         // Create log entry
         CreateLogMessagePara2 ( Timestamp   := SystemTime,
                                 MessageType := MessageType.CMD,
                                 Severity    := Severity.DEBUG,
                                 MessageCode := 0,
                                 MessageText := 'SyncSwLimits: Synchronization of SwLimits triggered by RC, SyncMode = {1}, SyncTime = {2}, SyncDirection = PLC -> RC',
                                 Para1       :=  SYNC_MODE_TO_STRING(AxesGroup.Parameter.Plc.Parameter.SynchronizationModes.SWLimits[SyncTime.AFTER_START_UP]),
                                 Para2       :=  SYNC_TIME_TO_STRING(SyncTime.AFTER_START_UP));
                                 RETURN;
			 END_IF
       
       // set timeout
       SetTimeout(PT := _rTimeout, rTimer := _rTimer);
       // jump back
      _rStep := 10;

       
  // ------------------------------------------
  // SyncMode : SERVER_TO_CLIENT 
  // ------------------------------------------
  12 : // Conflict triggerd by PLC ?  
       IF ( NOT AxesGroup.State.SyncStatePlc.InSync.SwLimits )
       THEN
         // set timeout
         SetTimeout(PT := _rTimeout, rTimer := _rTimer);
         // inc step counter
        _rStep := 20; // -> read RC data and write it to PLC                  

         // Create log entry
         CreateLogMessagePara2 ( Timestamp   := SystemTime,
                                 MessageType := MessageType.CMD,
                                 Severity    := Severity.DEBUG,
                                 MessageCode := 0,
                                 MessageText := 'SyncSwLimits: Synchronization of SwLimits triggered by PLC, SyncMode = {1}, SyncTime = {2}, SyncDirection = RC -> PLC',
                                 Para1       :=  SYNC_MODE_TO_STRING(AxesGroup.Parameter.Plc.Parameter.SynchronizationModes.SWLimits[SyncTime.AFTER_START_UP]),
                                 Para2       :=  SYNC_TIME_TO_STRING(SyncTime.AFTER_START_UP));
                                 RETURN;
       END_IF
   
       // Conflict triggered by RC ?
       IF ( NOT AxesGroup.State.SyncStateRc.InSync.SwLimits )
       THEN
         // set timeout
         SetTimeout(PT := _rTimeout, rTimer := _rTimer);
         // inc step counter
        _rStep := 20; // -> read RC data and write it to PLC

         // Create log entry
         CreateLogMessagePara2 ( Timestamp   := SystemTime,
                                 MessageType := MessageType.CMD,
                                 Severity    := Severity.DEBUG,
                                 MessageCode := 0,
                                 MessageText := 'SyncSwLimits: Synchronization of SwLimits triggered by RC, SyncMode = {1}, SyncTime = {2}, SyncDirection = RC -> PLC',
                                 Para1       :=  SYNC_MODE_TO_STRING(AxesGroup.Parameter.Plc.Parameter.SynchronizationModes.SWLimits[SyncTime.AFTER_START_UP]),
                                 Para2       :=  SYNC_TIME_TO_STRING(SyncTime.AFTER_START_UP));
                                 RETURN;
			 END_IF
       
       // set timeout
       SetTimeout(PT := _rTimeout, rTimer := _rTimer);
       // jump back
      _rStep := 10;
  

  // ------------------------------------------
  // SyncMode : AUTOMATIC 
  // ------------------------------------------
  13 : // Conflict triggerd by PLC ?  
       IF ( NOT AxesGroup.State.SyncStatePlc.InSync.SwLimits )
       THEN
         // set timeout
         SetTimeout(PT := _rTimeout, rTimer := _rTimer);
         // inc step counter
        _rStep := 30; // -> write PLC data to RC                  
         
         // Create log entry
         CreateLogMessagePara2 ( Timestamp   := SystemTime,
                                 MessageType := MessageType.CMD,
                                 Severity    := Severity.DEBUG,
                                 MessageCode := 0,
                                 MessageText := 'SyncSwLimits: Synchronization of SwLimits triggered by PLC, SyncMode = {1}, SyncTime = {2}, SyncDirection = PLC -> RC',
                                 Para1       :=  SYNC_MODE_TO_STRING(AxesGroup.Parameter.Plc.Parameter.SynchronizationModes.SWLimits[SyncTime.AFTER_START_UP]),
                                 Para2       :=  SYNC_TIME_TO_STRING(SyncTime.AFTER_START_UP));
                                 RETURN;
       END_IF
   
       // Conflict triggered by RC ?
       IF ( NOT AxesGroup.State.SyncStateRc.InSync.SwLimits )
       THEN
         // set timeout
         SetTimeout(PT := _rTimeout, rTimer := _rTimer);
         // inc step counter
        _rStep := 20; // -> read RC data an write it to PLC

         // Create log entry
         CreateLogMessagePara2 ( Timestamp   := SystemTime,
                                 MessageType := MessageType.CMD,
                                 Severity    := Severity.DEBUG,
                                 MessageCode := 0,
                                 MessageText := 'SyncSwLimits: Synchronization of SwLimits triggered by RC, SyncMode = {1}, SyncTime = {2}, SyncDirection = RC -> PLC',
                                 Para1       :=  SYNC_MODE_TO_STRING(AxesGroup.Parameter.Plc.Parameter.SynchronizationModes.SWLimits[SyncTime.AFTER_START_UP]),
                                 Para2       :=  SYNC_TIME_TO_STRING(SyncTime.AFTER_START_UP));
                                 RETURN;
			 END_IF
       
       // set timeout
       SetTimeout(PT := _rTimeout, rTimer := _rTimer);
       // jump back
      _rStep := 10; // ST-FIX F95: was commented out


  // ------------------------------------------
  // Read Data from RC and write it to PLC
  // ------------------------------------------
  20 : IF (( NOT _readRobotSWLimits.Busy  ) AND 
           ( NOT _readRobotSWLimits.Error ))
       THEN
         // execute command
        _readRobotSWLimits.Execute := TRUE;
         // set timeout
         SetTimeout(PT := _rTimeout, rTimer := _rTimer);
         // inc step counter
        _rStep := _rStep + 1;
       ELSE
         // check error ? 
         IF (_readRobotSWLimits.Error)
         THEN
           ErrorID     := _readRobotSWLimits.ErrorID;
           ErrorAddTxt := _readRobotSWLimits.ErrorAddTxt;
         END_IF  
       
         // timeout exceeded ? 
         IF (CheckTimeout(_rTimer) = RobotLibraryConstants.OK)
         THEN
           ErrorID     := RobotLibraryErrorIdEnum.ERR_TIMEOUT_CMD;
           ErrorAddTxt := CONCAT(_stepName, DINT_TO_STRING(_rStep));
         END_IF
       END_IF
 
  21 : IF (( NOT _readRobotSWLimits.Busy  ) AND
           ( NOT _readRobotSWLimits.Error ) AND
           (     _readRobotSWLimits.Done  ))
       THEN
         // reset execution
        _readRobotSWLimits.Execute := FALSE;
         // ST-FIX F107: AUTOMATIC - the PLC data were changed while the RC data were read: the PLC
         // change is the most recent one and is written to the RC instead of being overwritten
         IF ( AxesGroup.Parameter.Plc.Parameter.SynchronizationModes.SWLimits[SyncTime.AFTER_START_UP] = SyncMode.AUTOMATIC ) AND
            ( NOT IsSwLimitsEqual( Data1 := SwLimits, Data2 := _swLimits, IgnoreTimestamp := TRUE ))
         THEN
           // set timeout
           SetTimeout(PT := _rTimeout, rTimer := _rTimer);
           // -> write PLC data to RC
          _rStep := 30;
           RETURN;
         END_IF
         // update internal SwLimits data
         SwLimits := _readRobotSWLimits.OutCmd.LimitValues;         
        _swLimits := _readRobotSWLimits.OutCmd.LimitValues;
         // set timeout
         SetTimeout(PT := _rTimeout, rTimer := _rTimer);
         // inc step counter
        // ST-FIX F20: write the RC data back to reset DataChanged on the RC (spec 5.6.7.4.2)
        IF ( AxesGroup.State.RobotData.RCSupportedFunctions.WriteRobotSWLimits )
        THEN
          _rStep := 30;
        ELSE
          _rStep := 10;
        END_IF // -> jump to after startup           
       ELSE
         // check error ? 
         IF (_readRobotSWLimits.Error)
         THEN
           ErrorID     := _readRobotSWLimits.ErrorID;
           ErrorAddTxt := _readRobotSWLimits.ErrorAddTxt;           
         END_IF  
       
         // timeout exceeded ? 
         IF (CheckTimeout(_rTimer) = RobotLibraryConstants.OK)
         THEN
           ErrorID     := RobotLibraryErrorIdEnum.ERR_TIMEOUT_CMD;
           ErrorAddTxt := CONCAT(_stepName, DINT_TO_STRING(_rStep));
         END_IF
       END_IF


  // ------------------------------------------
  // Write data from PLC to RC
  // ------------------------------------------
  30 : IF (( NOT _writeRobotSWLimits.Busy  ) AND 
           ( NOT _writeRobotSWLimits.Error ))
       THEN
         // set command parameter
        _writeRobotSWLimits.ParCmd.ResetToFactoryDefaults := FALSE;      
        _writeRobotSWLimits.ParCmd.LimitValues :=  SwLimits;
         // execute command
        _writeRobotSWLimits.Execute := TRUE;
         // set timeout
         SetTimeout(PT := _rTimeout, rTimer := _rTimer);
         // inc step counter
        _rStep := _rStep + 1;
       ELSE
         // check error ? 
         IF (_writeRobotSWLimits.Error)
         THEN
           ErrorID     := _writeRobotSWLimits.ErrorID;
           ErrorAddTxt := _writeRobotSWLimits.ErrorAddTxt;;
         END_IF  
       
         // timeout exceeded ? 
         IF (CheckTimeout(_rTimer) = RobotLibraryConstants.OK)
         THEN
           ErrorID     := RobotLibraryErrorIdEnum.ERR_TIMEOUT_CMD;
           ErrorAddTxt := CONCAT(_stepName, DINT_TO_STRING(_rStep));
         END_IF
       END_IF
 
  31 : IF (( NOT _writeRobotSWLimits.Busy  ) AND
           ( NOT _writeRobotSWLimits.Error ) AND
           (     _writeRobotSWLimits.Done  ))
       THEN
         // execute command
        _writeRobotSWLimits.Execute := FALSE;      
         // update internal SwLimits data
        _swLimits := SwLimits; 
         // set timeout
         SetTimeout(PT := _rTimeout, rTimer := _rTimer);
         // inc step counter
        _rStep := 10; // -> jump to after startup;           
       ELSE
         // check error ? 
         IF (_writeRobotSWLimits.Error)
         THEN
           SetWarning( WarningID := RobotLibraryWarningIdEnum.WARN_SW_LIMITS_SYNC_FAILED_BY_ERROR_OF_READ_OR_WRITE_CMD, Overwrite := TRUE);    
         END_IF  
       
         // timeout exceeded ? 
         IF (CheckTimeout(_rTimer) = RobotLibraryConstants.OK)
         THEN
           ErrorID     := RobotLibraryErrorIdEnum.ERR_TIMEOUT_CMD;
           ErrorAddTxt := CONCAT(_stepName, DINT_TO_STRING(_rStep));
         END_IF
       END_IF
       
ELSE
  // invalid step
  ErrorID     := RobotLibraryErrorIdEnum.ERR_INVALID_STEP;
  ErrorAddTxt := CONCAT(_stepName , DINT_TO_STRING(_stepCmd));
END_CASE
END_METHOD

METHOD PRIVATE HandleSyncToolData
VAR_IN_OUT
   /// Robot assignment of function
  AxesGroup : AxesGroup;
  /// ToolData stored on PLC.For more information refer to 5.5.6.4
  ToolData  : ARRAY[*] OF Tool;
END_VAR 

VAR
  /// Internal step counter name
 _stepName        : STRING;    
  /// Internal reference to step counter
 _rStep           : REFERENCE TO DINT;
  /// Internal reference to timer
 _rTimer          : REFERENCE TO TON;
  /// Internal reference to timeout
 _rTimeout        : REFERENCE TO TIME; 
  /// Internal reference to synchroniztion index
 _rSyncIdx        : REFERENCE TO USINT;
  /// internal bit for condition found
 _found           : BOOL;
  /// empty data set to reset all DataChanged bits
 _dataChangedNone : AxesGroupStateDataChanged; 
  /// internal index for loops
 _idx             : DINT;
END_VAR
// Set internal references 
_stepName      :=   '_stepSyncToolData = ';
_rStep       REF=    _stepSyncToolData;
_rTimer      REF=   _timerSyncToolData;
_rTimeout    REF= _timeoutSyncToolData;
_rSyncIdx    REF=     _syncIdxToolData;


CASE _rStep
OF    
  0: // Check initialisation configured ?
     // ST-FIX F130: an invalid sync mode (warning of CheckParameterValid) -> no synchronization of the data set
     IF ((( _parCfg.PLC.Parameter.SynchronizationModes.Tool[SyncTime.DURING_START_UP] = SyncMode.NO_SYNCHRONIZATION ) AND
          ( _parCfg.PLC.Parameter.SynchronizationModes.Tool[SyncTime. AFTER_START_UP] = SyncMode.NO_SYNCHRONIZATION )) OR
         ( NOT SyncModesValid( During := _parCfg.PLC.Parameter.SynchronizationModes.Tool[SyncTime.DURING_START_UP],
                               After  := _parCfg.PLC.Parameter.SynchronizationModes.Tool[SyncTime. AFTER_START_UP] ) ))
     THEN
       RETURN;
     END_IF
     

     // wait for initialisation done
     IF  ((     AxesGroup.State.RobotData.RCSupportedFunctions. ReadToolData ) AND
          (     AxesGroup.State.RobotData.RCSupportedFunctions.WriteToolData ) AND
          (     AxesGroup.State.Initialized                                  ) AND 
          ( NOT Error                                                        ))  
     THEN
       // ST-FIX F102: count check after the initialization (HighestXIndex of this connection)
     // Check More Data on RC than on PLC -> Synchronization not possible
     IF (AxesGroup.State.ConfigurationData.HighestToolIndex > AxesGroup.SystemData.ToolDataCount)
     THEN
       SetError( ErrorID := RobotLibraryErrorIdEnum.ERR_SYNC_TOOL_COUNT_RC_HIGHER_THAN_PLC, Overwrite := FALSE);
       RETURN;
		 END_IF
       // Check PLC tools < RC tools and SyncTool enabled ?    
       IF (( AxesGroup.State.DataEnableSync.EnableSyncTool      = TRUE                             )  AND
           ( AxesGroup.Parameter.Rob.Parameter.HighestToolIndex > AxesGroup.SystemData.ToolDataMax ))        
       THEN
         SetWarning( WarningID := RobotLibraryWarningIdEnum.WARN_TOOL_DATA_ARRAY_TOO_SHORT, Overwrite := TRUE);
       END_IF

       // Create log entry
       CreateLogMessagePara1 ( Timestamp   := SystemTime,
                               MessageType := MessageType.CMD,
                               Severity    := Severity.DEBUG,
                               MessageCode := 0,
                               MessageText := 'SyncToolData: Start initial reading of ToolData from RC',
                               Para1       :=  '');
       
       // init tool number
      _rSyncIdx := LIMIT(1, DINT_TO_USINT(AxesGroup.SystemData.ToolDataMin), AxesGroup.State.UnifiedToolIndex); // ST-FIX F21: index 0 is fixed on the RC 
       // init count of unsynchronized elements
       AxesGroup.State.SyncStatePlc.UnSyncNo.Tool := 0;
       // set timeout
       SetTimeout(PT := _rTimeout, rTimer := _rTimer);
       // inc step counter
      _rStep := _rStep + 1;
     END_IF     

     
     // Start read ToolData
  1: IF (( NOT _readToolData.Busy  ) AND 
         ( NOT _readToolData.Error ) AND
         ( NOT _readToolData.Done  ))
     THEN
       // set command parameter
      _readToolData.ParCmd.ToolNo := _rSyncIdx;      
       // execute command
      _readToolData.Execute := TRUE;
       // set timeout
       SetTimeout(PT := _rTimeout, rTimer := _rTimer);
       // inc step counter
      _rStep := _rStep + 1;
     ELSE
       // check error ? 
       IF ( _readToolData.Error ) AND ( WarningID = RobotLibraryWarningIdEnum.NO_WARNING )
       THEN
         SetWarning( WarningID := RobotLibraryWarningIdEnum.WARN_TOOL_SYNC_FAILED_BY_ERROR_OF_READ_OR_WRITE_CMD, Overwrite := TRUE);           
       END_IF  
       
       // timeout exceeded ? 
       IF (CheckTimeout(_rTimer) = RobotLibraryConstants.OK)
       THEN
         ErrorID     := RobotLibraryErrorIdEnum.ERR_TIMEOUT_CMD;
         ErrorAddTxt := CONCAT(_stepName, DINT_TO_STRING(_rStep));
       END_IF
     END_IF
 
     
     // Wait Tooldata read
  2: IF (( NOT _readToolData.Busy  ) AND
         ( NOT _readToolData.Error ) AND
         (     _readToolData.Done  ))
     THEN
       // reset execution
      _readToolData.Execute := FALSE;
       // set available bit
      _toolData[_rSyncIdx].Available := TRUE; 
       ToolData[_rSyncIdx].Available := TRUE;      
       // Copy data
      _toolData[_rSyncIdx].Data := _readToolData.OutCmd.ToolData;

       // Check tool data is equal ? 
       IF ( NOT IsToolDataEqual( Data1 := _toolData[_rSyncIdx].Data, Data2 := ToolData[_rSyncIdx].Data, IgnoreTimestamp := TRUE))
       THEN
         // Reset plc in sync flag
         AxesGroup.State.SyncStatePlc.InSync.Tool := FALSE;
         // Set data changed flag
         AxesGroup.State.DataChanged.Tool[_rSyncIdx] := TRUE;
         // inc count of unsynchronised plc tools
         AxesGroup.State.SyncStatePlc.UnSyncNo.Tool := AxesGroup.State.SyncStatePlc.UnSyncNo.Tool + 1;
        
         // Create log entry
         CreateLogMessagePara1 ( Timestamp   := SystemTime,
                                 MessageType := MessageType.CMD,
                                 Severity    := Severity.DEBUG,
                                 MessageCode := 0,
                                 MessageText := 'SyncToolData: Detected a difference in Tool[{1}] between PLC and RC',
                                 Para1       :=  DINT_TO_STRING(_rSyncIdx));
        
        
         // Check synchronisation is enabled ? 
         IF ( NOT AxesGroup.State.DataEnableSync.EnableSyncTool ) AND (InfoID = RobotLibraryInfoIdEnum.NO_INFO )
         THEN
           SetInfo( InfoID := RobotLibraryInfoIdEnum.INFO_SYNC_TOOL_DATA_DISABLED, Overwrite := TRUE);
				 END_IF
         
         // Check user interaction needed ?  
         IF ( AxesGroup.Parameter.PLC.Parameter.SyncUserInteraction.Tool ) AND ( WarningID = RobotLibraryWarningIdEnum.NO_WARNING )
         THEN
           SetWarning( WarningID := RobotLibraryWarningIdEnum.WARN_TOOL_NUMBER_SYNC_ERROR, Overwrite :=  TRUE);                    
				 END_IF
			 END_IF
             
       // Check all tools read ? 
       IF ( _rSyncIdx < AxesGroup.State.UnifiedToolIndex )
       THEN
         // set timeout
         SetTimeout(PT := _rTimeout, rTimer := _rTimer);
         // inc tool index
        _rSyncIdx := _rSyncIdx + 1;
         // dec step counter
        _rStep := _rStep - 1;
       ELSE
         // set timeout
         SetTimeout(PT := _rTimeout, rTimer := _rTimer);
         // inc step counter
        _rStep := _rStep + 1;           
       END_IF
     ELSE
       // check error ? 
       IF (_readToolData.Error)
       THEN
         // Set warning
         SetWarning( WarningID := RobotLibraryWarningIdEnum.WARN_TOOL_SYNC_FAILED_BY_ERROR_OF_READ_OR_WRITE_CMD, Overwrite := TRUE);                    
         // reset available bit
         ToolData[_rSyncIdx].Available := FALSE;
        _toolData[_rSyncIdx].Available := FALSE;
       END_IF  
       
       // timeout exceeded ? 
       IF (CheckTimeout(_rTimer) = RobotLibraryConstants.OK)
       THEN
         ErrorID     := RobotLibraryErrorIdEnum.ERR_TIMEOUT_CMD;
         ErrorAddTxt := CONCAT(_stepName, DINT_TO_STRING(_rStep));
       END_IF
     END_IF
     
     
     // Check synchronisation state ? 
  3: IF (( AxesGroup.State.SyncStatePlc.UnSyncNo.Tool                                            = 0                           ) OR 
         ( AxesGroup.Parameter.Plc.Parameter.SynchronizationModes.Tool[SyncTime.DURING_START_UP] = SyncMode.NO_SYNCHRONIZATION ))
     THEN
       // Update bit for data in sync
       AxesGroup.State.SyncStatePlc.InSync.Tool := (AxesGroup.State.SyncStatePlc.UnSyncNo.Tool = 0);
         // ST-FIX F165: synchronization of the start-up phase finished
         AxesGroup.State.Synchronizing.Tool := FALSE;
       // set timeout
       SetTimeout(PT := _rTimeout, rTimer := _rTimer);
       // inc step counter
      _rStep := 10; // -> jump to after startup
            
       // Create log entry
       CreateLogMessagePara1 ( Timestamp   := SystemTime,
                               MessageType := MessageType.CMD,
                               Severity    := Severity.DEBUG,
                               MessageCode := 0,
                               MessageText := 'SyncToolData: Synchronization Startup Phase done',
                               Para1       :=  '' );      
     ELSE 
       // Check user interaction needed ? 
       IF ( NOT AxesGroup.Parameter.PLC.Parameter.SyncUserInteraction.Tool )
       THEN
         CASE AxesGroup.Parameter.Plc.Parameter.SynchronizationModes.Tool[SyncTime.DURING_START_UP] OF

           SyncMode.SERVER_TO_CLIENT : 

           
             FOR _idx := AxesGroup.SystemData.ToolDataMin TO MIN(AxesGroup.SystemData.ToolDataMax, RobotLibraryParameter.TOOL_MAX - 1) // ST-FIX F18
             DO
               // Overwrite PLC data with RC data
               ToolData[_idx] := _toolData[_idx];            
						 END_FOR
             // Reset data changed flags
             AxesGroup.State.DataChanged.Tool := _dataChangedNone.Tool;
             // Reset Synchronizing flag
             AxesGroup.State.Synchronizing.Tool := FALSE;
             // Set plc in sync flag
             AxesGroup.State.SyncStatePlc.InSync.Tool := TRUE;
             // Reset count of unsynchronised plc tools
             AxesGroup.State.SyncStatePlc.UnSyncNo.Tool := 0;            
             // set timeout
             SetTimeout(PT := _rTimeout, rTimer := _rTimer);
             // inc step counter
            _rStep := 10; // -> jump to after startup         

            // Create log entry
            CreateLogMessagePara3 ( Timestamp   := SystemTime,
                                    MessageType := MessageType.CMD,
                                    Severity    := Severity.DEBUG,
                                    MessageCode := 0,
                                    MessageText := 'SyncToolData: Synchronization of Tools triggered by StartUp-Compare, SyncMode = {2}, SyncTime = {3}, SyncDirection = RC -> PLC',
                                    Para1       :=  DINT_TO_STRING(_rSyncIdx),
                                    Para2       :=  SYNC_MODE_TO_STRING(AxesGroup.Parameter.Plc.Parameter.SynchronizationModes.Tool[SyncTime.DURING_START_UP]),
                                    Para3       :=  SYNC_TIME_TO_STRING(SyncTime.DURING_START_UP));
            // Create log entry
            CreateLogMessagePara1 ( Timestamp   := SystemTime,
                                    MessageType := MessageType.CMD,
                                    Severity    := Severity.DEBUG,
                                    MessageCode := 0,
                                    MessageText := 'SyncToolData: Applied the initial read tool data from RC',
                                    Para1       :=  '' );

				   SyncMode.CLIENT_TO_SERVER : ;

             // Check conflicts to solve ? 
             FOR _rSyncIdx := 1 TO AxesGroup.State.UnifiedToolIndex // ST-FIX F21: index 0 is fixed on the RC
             DO
               IF ( AxesGroup.State.DataChanged.Tool[_rSyncIdx] )
               THEN
                _found := TRUE;
                 EXIT;
		  			   END_IF
             END_FOR
           
             IF ( _found ) 
             THEN
               // Reset plc in sync flag
               AxesGroup.State.SyncStatePlc.InSync.Tool := FALSE;
               // Set Synchronizing flag
               AxesGroup.State.Synchronizing.Tool := TRUE;
               // set timeout
               SetTimeout(PT := _rTimeout, rTimer := _rTimer);
               // inc step counter
              _rStep := _rStep +1; // -> write PLC data to RC                  
               // Create log entry
               CreateLogMessagePara3 ( Timestamp   := SystemTime,
                                       MessageType := MessageType.CMD,
                                       Severity    := Severity.DEBUG,
                                       MessageCode := 0,
                                       MessageText := 'SyncToolData: Synchronization of Tool[{1}] triggered by StartUp-Compare, SyncMode = {2}, SyncTime = {3}, SyncDirection = PLC -> RC',
                                       Para1       :=  DINT_TO_STRING(_rSyncIdx),
                                       Para2       :=  SYNC_MODE_TO_STRING(AxesGroup.Parameter.Plc.Parameter.SynchronizationModes.Tool[SyncTime.DURING_START_UP]),
                                       Para3       :=  SYNC_TIME_TO_STRING(SyncTime.DURING_START_UP));
             ELSE
               // Reset data changed flags
               AxesGroup.State.DataChanged.Tool := _dataChangedNone.Tool;
               // Reset Synchronizing flag
               AxesGroup.State.Synchronizing.Tool := FALSE;
               // Set plc in sync flag
               AxesGroup.State.SyncStatePlc.InSync.Tool := TRUE;
               // Reset count of unsynchronised tools
               AxesGroup.State.SyncStatePlc.UnSyncNo.Tool := 0;
               // set timeout
               SetTimeout(PT := _rTimeout, rTimer := _rTimer);
               // inc step counter
              _rStep := 10; // -> jump to after startup                  
				     END_IF
         ELSE
           // invalid sync mode for startup
           SetWarning( WarningID := RobotLibraryWarningIdEnum.WARN_TOOL_DATA_SYNC_MODE_INVALID, Overwrite := TRUE ); // ST-FIX F130: warning instead of the own error
 	       END_CASE
       ELSE
         // ST-FIX F94: the user resolves the conflict with the write / read functions - read the RC data again
         IF ( CheckTimeout(_rTimer) = RobotLibraryConstants.OK )
         THEN
           AxesGroup.State.DataChanged.Tool := _dataChangedNone.Tool;
           SetTimeout(PT := _rTimeout, rTimer := _rTimer);
          _rStep := 0; // -> read the RC data and compare again
         END_IF
       END_IF
     END_IF  

     
     // Start write tool data  
  4: IF (( NOT _writeToolData.Busy  ) AND 
         ( NOT _writeToolData.Error ))
     THEN
       // set command parameter
      _writeToolData.ParCmd.ToolNo   := _rSyncIdx;      
      _writeToolData.ParCmd.ToolData :=  ToolData[_rSyncIdx].Data;
       // execute command
      _writeToolData.Execute := TRUE;
       // set timeout
       SetTimeout(PT := _rTimeout, rTimer := _rTimer);
       // inc step counter
      _rStep := _rStep + 1;
     ELSE
       // check error ? 
       IF (_writeToolData.Error)
       THEN
         ErrorID     := _writeToolData.ErrorID;
         ErrorAddTxt := _writeToolData.ErrorAddTxt;;
       END_IF  
       
       // timeout exceeded ? 
       IF (CheckTimeout(_rTimer) = RobotLibraryConstants.OK)
       THEN
         ErrorID     := RobotLibraryErrorIdEnum.ERR_TIMEOUT_CMD;
         ErrorAddTxt := CONCAT(_stepName, DINT_TO_STRING(_rStep));
       END_IF
     END_IF
 
     
     // Wait tool data written ?   
  5: IF (( NOT _writeToolData.Busy  ) AND
         ( NOT _writeToolData.Error ) AND
         (     _writeToolData.Done  ))
     THEN
       // execute command
      _writeToolData.Execute := FALSE;
       // apply tool data to internal tool data
      _toolData[_rSyncIdx] := ToolData[_rSyncIdx];
       // reset data changed bit 
       AxesGroup.State.DataChanged.Tool[_rSyncIdx] := FALSE;
       // dec count of unsynchronised tools
       AxesGroup.State.SyncStatePlc.UnSyncNo.Tool := AxesGroup.State.SyncStatePlc.UnSyncNo.Tool - 1;
       // set timeout        
       SetTimeout(PT := _rTimeout, rTimer := _rTimer);
       // dec step counter
      _rStep := _rStep - 2; 
     ELSE
       // check error ? 
       IF (_writeToolData.Error)
       THEN
         SetWarning( WarningID := RobotLibraryWarningIdEnum.WARN_TOOL_SYNC_FAILED_BY_ERROR_OF_READ_OR_WRITE_CMD, Overwrite := TRUE);
           // ST-FIX F168: refused by the RC -> warning, go on with the next entry
          _writeToolData.Execute := FALSE;
          _toolData[_rSyncIdx] := ToolData[_rSyncIdx];
          AxesGroup.State.DataChanged.Tool[_rSyncIdx] := FALSE;
          AxesGroup.State.SyncStatePlc.UnSyncNo.Tool := AxesGroup.State.SyncStatePlc.UnSyncNo.Tool - 1;
           SetTimeout(PT := _rTimeout, rTimer := _rTimer);
          _rStep := _rStep - 2;           
       END_IF  
       
       // timeout exceeded ? 
       IF (CheckTimeout(_rTimer) = RobotLibraryConstants.OK)
       THEN
         ErrorID     := RobotLibraryErrorIdEnum.ERR_TIMEOUT_CMD;
         ErrorAddTxt := CONCAT(_stepName, DINT_TO_STRING(_rStep));
       END_IF
     END_IF

     
  // --------------------------------------------
  // SyncMode after startup : 
  // --------------------------------------------
         
  10 :// check synchronisation active ? 
       // ST-FIX F93: compare also with NO_SYNCHRONIZATION (no transfer, see the CASE below)

       // reset count of unsynchronised tools
       AxesGroup.State.SyncStatePlc.UnSyncNo.Tool := 0;

       // Check all tool datas
       FOR _rSyncIdx := 1 TO AxesGroup.State.UnifiedToolIndex // ST-FIX F21: index 0 is fixed on the RC
       DO
         // compare tool data
         AxesGroup.State.DataChanged.Tool[_rSyncIdx] := NOT IsToolDataEqual( Data1 := ToolData[_rSyncIdx].Data, Data2 := _toolData[_rSyncIdx].Data, IgnoreTimestamp := TRUE (* ST-FIX F57 *));

         // Check Tool data changed ? 
         IF (AxesGroup.State.DataChanged.Tool[_rSyncIdx])
         THEN
           // inc count of unsynchronised plc tools
           AxesGroup.State.SyncStatePlc.UnSyncNo.Tool := AxesGroup.State.SyncStatePlc.UnSyncNo.Tool + 1;
           // Create log entry
           CreateLogMessagePara2 ( Timestamp   := SystemTime,
                                   MessageType := MessageType.CMD,
                                   Severity    := Severity.DEBUG,
                                   MessageCode := 0,
                                   MessageText := 'SyncToolData: Detected a local change of Tool[{1}] on PLC, SyncTime = {2}',
                                   Para1       :=  DINT_TO_STRING(_rSyncIdx),    
                                   Para2       :=  SYNC_TIME_TO_STRING(SyncTime.AFTER_START_UP));       
				 END_IF

         // Update plc in sync flag
         AxesGroup.State.SyncStatePlc.InSync.Tool := (AxesGroup.State.SyncStatePlc.UnSyncNo.Tool = 0); 
	     END_FOR

       // Check synchronization is needed ? 
       IF ( NOT AxesGroup.State.SyncStatePlc.InSync.Tool ) XOR  
          ( NOT AxesGroup.State.SyncStateRc .InSync.Tool )
       THEN
         CASE AxesGroup.Parameter.Plc.Parameter.SynchronizationModes.Tool[SyncTime.AFTER_START_UP] 
         OF         
           // NO_SYNCHRONIZATION
           SyncMode.NO_SYNCHRONIZATION : ; // no further action 
           
           // CLIENT_TO_SERVER
           SyncMode.CLIENT_TO_SERVER :
             // set timeout
             SetTimeout(PT := _rTimeout, rTimer := _rTimer);
             // inc step counter
            _rStep := 11;
  
           // SERVER_TO_CLIENT
           SyncMode.SERVER_TO_CLIENT :
             // set timeout
             SetTimeout(PT := _rTimeout, rTimer := _rTimer);
             // inc step counter
            _rStep := 12;
  
           // AUTOMATIC
           SyncMode.AUTOMATIC : 
             // set timeout
             SetTimeout(PT := _rTimeout, rTimer := _rTimer);
             // inc step counter
            _rStep := 13;
         END_CASE
       ELSE
         // datas changeḍ on both sides ? -> Warning 
         IF (( NOT AxesGroup.State.SyncStatePlc.InSync.Tool ) AND  
             ( NOT AxesGroup.State.SyncStateRc .InSync.Tool ))
         THEN
           // ST-FIX F58: CLIENT_TO_SERVER / SERVER_TO_CLIENT decide the direction also if both sides changed
CASE AxesGroup.Parameter.Plc.Parameter.SynchronizationModes.Tool[SyncTime.AFTER_START_UP] OF
  SyncMode.CLIENT_TO_SERVER : _rStep := 11;
  SyncMode.SERVER_TO_CLIENT : _rStep := 12;
ELSE
  SetWarning( WarningID := RobotLibraryWarningIdEnum.WARN_TOOL_SYNC_BOTH_SIDES_CHANGED, Overwrite := TRUE);
END_CASE
         END_IF
       END_IF


  // ------------------------------------------
  // SyncMode : CLIENT_TO_SERVER 
  // ------------------------------------------  
  11 : // Conflict triggerd by PLC ?  
       IF ( NOT AxesGroup.State.SyncStatePlc.InSync.Tool )
       THEN
         // search for changed index  
         FOR _rSyncIdx := 1 TO AxesGroup.State.UnifiedToolIndex // ST-FIX F21: index 0 is fixed on the RC
         DO
           IF ( AxesGroup.State.DataChanged.Tool[_rSyncIdx] )
           THEN
             // set timeout
             SetTimeout(PT := _rTimeout, rTimer := _rTimer);
             // inc step counter
            _rStep := 30; // -> write PLC data to RC                  
             EXIT;             
					 END_IF
         END_FOR
         
         // Create log entry
         CreateLogMessagePara3 ( Timestamp   := SystemTime,
                                 MessageType := MessageType.CMD,
                                 Severity    := Severity.DEBUG,
                                 MessageCode := 0,
                                 MessageText := 'SyncToolData: Synchronization of Tool[{1}] triggered by PLC, SyncMode = {2}, SyncTime = {3}, SyncDirection = PLC -> RC',
                                 Para1       :=  DINT_TO_STRING(_rSyncIdx),
                                 Para2       :=  SYNC_MODE_TO_STRING(AxesGroup.Parameter.Plc.Parameter.SynchronizationModes.Tool[SyncTime.AFTER_START_UP]),
                                 Para3       :=  SYNC_TIME_TO_STRING(SyncTime.AFTER_START_UP));
                                 RETURN;
       END_IF
   
       // Conflict triggered by RC ?
       IF ( NOT AxesGroup.State.SyncStateRc.InSync.Tool )
       THEN
         // get changed index 
        _rSyncIdx :=  LIMIT(1, AxesGroup.State.SyncStateRc.UnSyncNo.Tool, // ST-FIX F21: index 0 is fixed on the RC
 AxesGroup.State.UnifiedToolIndex);
         // set timeout
         SetTimeout(PT := _rTimeout, rTimer := _rTimer);
         // inc step counter
        _rStep := 30; // -> write PLC data to RC

         // Create log entry
         CreateLogMessagePara3 ( Timestamp   := SystemTime,
                                 MessageType := MessageType.CMD,
                                 Severity    := Severity.DEBUG,
                                 MessageCode := 0,
                                 MessageText := 'SyncToolData: Synchronization of Tool[{1}] triggered by RC, SyncMode = {2}, SyncTime = {3}, SyncDirection = PLC -> RC',
                                 Para1       :=  DINT_TO_STRING(_rSyncIdx),
                                 Para2       :=  SYNC_MODE_TO_STRING(AxesGroup.Parameter.Plc.Parameter.SynchronizationModes.Tool[SyncTime.AFTER_START_UP]),
                                 Para3       :=  SYNC_TIME_TO_STRING(SyncTime.AFTER_START_UP));
                                 RETURN;
			 END_IF
       
       // set timeout
       SetTimeout(PT := _rTimeout, rTimer := _rTimer);
       // jump back
      _rStep := 10;

       
  // ------------------------------------------
  // SyncMode : SERVER_TO_CLIENT 
  // ------------------------------------------
  12 : // Conflict triggerd by PLC ?  
       IF ( NOT AxesGroup.State.SyncStatePlc.InSync.Tool )
       THEN
         // search for changed index  
         FOR _rSyncIdx := 1 TO AxesGroup.State.UnifiedToolIndex // ST-FIX F21: index 0 is fixed on the RC
         DO
           IF ( AxesGroup.State.DataChanged.Tool[_rSyncIdx] )
           THEN
             // set timeout
             SetTimeout(PT := _rTimeout, rTimer := _rTimer);
             // inc step counter
            _rStep := 20; // -> read RC data and write it to PLC                  
             EXIT;
					 END_IF
         END_FOR

         // Create log entry
         CreateLogMessagePara3 ( Timestamp   := SystemTime,
                                 MessageType := MessageType.CMD,
                                 Severity    := Severity.DEBUG,
                                 MessageCode := 0,
                                 MessageText := 'SyncToolData: Synchronization of Tool[{1}] triggered by PLC, SyncMode = {2}, SyncTime = {3}, SyncDirection = RC -> PLC',
                                 Para1       :=  DINT_TO_STRING(_rSyncIdx),
                                 Para2       :=  SYNC_MODE_TO_STRING(AxesGroup.Parameter.Plc.Parameter.SynchronizationModes.Tool[SyncTime.AFTER_START_UP]),
                                 Para3       :=  SYNC_TIME_TO_STRING(SyncTime.AFTER_START_UP));
                                 RETURN;
       END_IF
   
       // Conflict triggered by RC ?
       IF ( NOT AxesGroup.State.SyncStateRc.InSync.Tool )
       THEN
         // get changed index 
        _rSyncIdx := LIMIT(1, AxesGroup.State.SyncStateRc.UnSyncNo.Tool, // ST-FIX F21: index 0 is fixed on the RC
 AxesGroup.State.UnifiedToolIndex);
         // set timeout
         SetTimeout(PT := _rTimeout, rTimer := _rTimer);
         // inc step counter
        _rStep := 20; // -> read RC data and write it to PLC

         // Create log entry
         CreateLogMessagePara3 ( Timestamp   := SystemTime,
                                 MessageType := MessageType.CMD,
                                 Severity    := Severity.DEBUG,
                                 MessageCode := 0,
                                 MessageText := 'SyncToolData: Synchronization of Tool[{1}] triggered by RC, SyncMode = {2}, SyncTime = {3}, SyncDirection = RC -> PLC',
                                 Para1       :=  DINT_TO_STRING(_rSyncIdx),
                                 Para2       :=  SYNC_MODE_TO_STRING(AxesGroup.Parameter.Plc.Parameter.SynchronizationModes.Tool[SyncTime.AFTER_START_UP]),
                                 Para3       :=  SYNC_TIME_TO_STRING(SyncTime.AFTER_START_UP));
                                 RETURN;
			 END_IF
       
       // set timeout
       SetTimeout(PT := _rTimeout, rTimer := _rTimer);
       // jump back
      _rStep := 10;
  

  // ------------------------------------------
  // SyncMode : AUTOMATIC 
  // ------------------------------------------
  13 : // Conflict triggerd by PLC ?  
       IF ( NOT AxesGroup.State.SyncStatePlc.InSync.Tool )
       THEN
         // search for changed index  
         FOR _rSyncIdx := 1 TO AxesGroup.State.UnifiedToolIndex // ST-FIX F21: index 0 is fixed on the RC
         DO
           IF ( AxesGroup.State.DataChanged.Tool[_rSyncIdx] )
           THEN
             // set timeout
             SetTimeout(PT := _rTimeout, rTimer := _rTimer);
             // inc step counter
            _rStep := 30; // -> write PLC data to RC                  
             EXIT;
					 END_IF
         END_FOR
         
         // Create log entry
         CreateLogMessagePara3 ( Timestamp   := SystemTime,
                                 MessageType := MessageType.CMD,
                                 Severity    := Severity.DEBUG,
                                 MessageCode := 0,
                                 MessageText := 'SyncToolData: Synchronization of Tool[{1}] triggered by PLC, SyncMode = {2}, SyncTime = {3}, SyncDirection = PLC -> RC',
                                 Para1       :=  DINT_TO_STRING(_rSyncIdx),
                                 Para2       :=  SYNC_MODE_TO_STRING(AxesGroup.Parameter.Plc.Parameter.SynchronizationModes.Tool[SyncTime.AFTER_START_UP]),
                                 Para3       :=  SYNC_TIME_TO_STRING(SyncTime.AFTER_START_UP));
                                 RETURN;
       END_IF
   
       // Conflict triggered by RC ?
       IF ( NOT AxesGroup.State.SyncStateRc.InSync.Tool )
       THEN
         // get changed index 
        _rSyncIdx := LIMIT(1, AxesGroup.State.SyncStateRc.UnSyncNo.Tool, // ST-FIX F21: index 0 is fixed on the RC
 AxesGroup.State.UnifiedToolIndex);
         // set timeout
         SetTimeout(PT := _rTimeout, rTimer := _rTimer);
         // inc step counter
        _rStep := 20; // -> read RC data an write it to PLC

         // Create log entry
         CreateLogMessagePara3 ( Timestamp   := SystemTime,
                                 MessageType := MessageType.CMD,
                                 Severity    := Severity.DEBUG,
                                 MessageCode := 0,
                                 MessageText := 'SyncToolData: Synchronization of Tool[{1}] triggered by RC, SyncMode = {2}, SyncTime = {3}, SyncDirection = RC -> PLC',
                                 Para1       :=  DINT_TO_STRING(_rSyncIdx),
                                 Para2       :=  SYNC_MODE_TO_STRING(AxesGroup.Parameter.Plc.Parameter.SynchronizationModes.Tool[SyncTime.AFTER_START_UP]),
                                 Para3       :=  SYNC_TIME_TO_STRING(SyncTime.AFTER_START_UP));
                                 RETURN;
			 END_IF
       
       // set timeout
       SetTimeout(PT := _rTimeout, rTimer := _rTimer);
       // jump back
      _rStep := 10; // ST-FIX F95: was commented out


  // ------------------------------------------
  // Read Data from RC and write it to PLC
  // ------------------------------------------
  20 : IF (( NOT _readToolData.Busy  ) AND 
           ( NOT _readToolData.Error ))
       THEN
         // set command parameter
        _readToolData.ParCmd.ToolNo := _rSyncIdx;      
         // execute command
        _readToolData.Execute := TRUE;
         // set timeout
         SetTimeout(PT := _rTimeout, rTimer := _rTimer);
         // inc step counter
        _rStep := _rStep + 1;
       ELSE
         // check error ? 
         IF (_readToolData.Error)
         THEN
           ErrorID     := _readToolData.ErrorID;
           ErrorAddTxt := _readToolData.ErrorAddTxt;
         END_IF  
       
         // timeout exceeded ? 
         IF (CheckTimeout(_rTimer) = RobotLibraryConstants.OK)
         THEN
           ErrorID     := RobotLibraryErrorIdEnum.ERR_TIMEOUT_CMD;
           ErrorAddTxt := CONCAT(_stepName, DINT_TO_STRING(_rStep));
         END_IF
       END_IF
 
  21 : IF (( NOT _readToolData.Busy  ) AND
           ( NOT _readToolData.Error ) AND
           (     _readToolData.Done  ))
       THEN
         // reset execution
        _readToolData.Execute := FALSE;
         // ST-FIX F107: AUTOMATIC - the PLC data were changed while the RC data were read: the PLC
         // change is the most recent one and is written to the RC instead of being overwritten
         IF ( AxesGroup.Parameter.Plc.Parameter.SynchronizationModes.Tool[SyncTime.AFTER_START_UP] = SyncMode.AUTOMATIC ) AND
            ( NOT IsToolDataEqual( Data1 := ToolData[_rSyncIdx].Data, Data2 := _toolData[_rSyncIdx].Data, IgnoreTimestamp := TRUE ))
         THEN
           // set timeout
           SetTimeout(PT := _rTimeout, rTimer := _rTimer);
           // -> write PLC data to RC
          _rStep := 30;
           RETURN;
         END_IF
         // update internal tool data
         ToolData[_rSyncIdx].Data := _readToolData.OutCmd.ToolData;         
        _toolData[_rSyncIdx].Data := _readToolData.OutCmd.ToolData;
         // set available bit
         ToolData[_rSyncIdx].Available := TRUE;
        _toolData[_rSyncIdx].Available := TRUE;
         // set timeout
         SetTimeout(PT := _rTimeout, rTimer := _rTimer);
         // inc step counter
        // ST-FIX F20: write the RC data back to reset DataChanged on the RC (spec 5.6.7.4.2)
        IF ( AxesGroup.State.RobotData.RCSupportedFunctions.WriteToolData )
        THEN
          _rStep := 30;
        ELSE
          _rStep := 10;
        END_IF // -> jump to after startup           
       ELSE
         // check error ? 
         IF (_readToolData.Error)
         THEN
           ErrorID     := _readToolData.ErrorID;
           ErrorAddTxt := _readToolData.ErrorAddTxt;           
           // reset available bit
           ToolData[_rSyncIdx].Available := FALSE;
          _toolData[_rSyncIdx].Available := FALSE;
         END_IF  
       
         // timeout exceeded ? 
         IF (CheckTimeout(_rTimer) = RobotLibraryConstants.OK)
         THEN
           ErrorID     := RobotLibraryErrorIdEnum.ERR_TIMEOUT_CMD;
           ErrorAddTxt := CONCAT(_stepName, DINT_TO_STRING(_rStep));
         END_IF
       END_IF


  // ------------------------------------------
  // Write data from PLC to RC
  // ------------------------------------------
  30 : IF (( NOT _writeToolData.Busy  ) AND 
           ( NOT _writeToolData.Error ))
       THEN
         // set command parameter
        _writeToolData.ParCmd.ToolNo   := _rSyncIdx;      
        _writeToolData.ParCmd.ToolData :=  ToolData[_rSyncIdx].Data;
         // execute command
        _writeToolData.Execute := TRUE;
         // set timeout
         SetTimeout(PT := _rTimeout, rTimer := _rTimer);
         // inc step counter
        _rStep := _rStep + 1;
       ELSE
         // check error ? 
         IF (_writeToolData.Error)
         THEN
           ErrorID     := _writeToolData.ErrorID;
           ErrorAddTxt := _writeToolData.ErrorAddTxt;;
         END_IF  
       
         // timeout exceeded ? 
         IF (CheckTimeout(_rTimer) = RobotLibraryConstants.OK)
         THEN
           ErrorID     := RobotLibraryErrorIdEnum.ERR_TIMEOUT_CMD;
           ErrorAddTxt := CONCAT(_stepName, DINT_TO_STRING(_rStep));
         END_IF
       END_IF
 
  31 : IF (( NOT _writeToolData.Busy  ) AND
           ( NOT _writeToolData.Error ) AND
           (     _writeToolData.Done  ))
       THEN
         // execute command
        _writeToolData.Execute := FALSE;      
         // update internal tool data
        _toolData[_rSyncIdx] := ToolData[_rSyncIdx]; 
         // set available bit
         ToolData[_rSyncIdx].Available := TRUE; 
        _toolData[_rSyncIdx].Available := TRUE;         
         // set timeout
         SetTimeout(PT := _rTimeout, rTimer := _rTimer);
         // inc step counter
        _rStep := 10; // -> jump to after startup;           
       ELSE
         // check error ? 
         IF (_writeToolData.Error)
         THEN
           SetWarning( WarningID := RobotLibraryWarningIdEnum.WARN_TOOL_SYNC_FAILED_BY_ERROR_OF_READ_OR_WRITE_CMD, Overwrite := TRUE);    
           // reset available bit
           ToolData[_rSyncIdx].Available := FALSE;
          _toolData[_rSyncIdx].Available := FALSE;
         END_IF  
       
         // timeout exceeded ? 
         IF (CheckTimeout(_rTimer) = RobotLibraryConstants.OK)
         THEN
           ErrorID     := RobotLibraryErrorIdEnum.ERR_TIMEOUT_CMD;
           ErrorAddTxt := CONCAT(_stepName, DINT_TO_STRING(_rStep));
         END_IF
       END_IF
       
ELSE
  // invalid step
  ErrorID     := RobotLibraryErrorIdEnum.ERR_INVALID_STEP;
  ErrorAddTxt := CONCAT(_stepName , DINT_TO_STRING(_stepCmd));
END_CASE
END_METHOD

METHOD PRIVATE HandleSyncWorkArea
VAR_IN_OUT
   /// Robot assignment of function
  AxesGroup : AxesGroup;
  /// Work areas stored on PLC. For more information refer to 5.5.8
  WorkAreas : ARRAY[*] OF RobotWorkArea;
END_VAR 

VAR
  /// Internal step counter name
 _stepName        : STRING;    
  /// Internal reference to step counter
 _rStep           : REFERENCE TO DINT;
  /// Internal reference to timer
 _rTimer          : REFERENCE TO TON;
  /// Internal reference to timeout
 _rTimeout        : REFERENCE TO TIME; 
  /// Internal reference to synchroniztion index
 _rSyncIdx        : REFERENCE TO USINT;
  /// internal bit for condition found
 _found           : BOOL;
  /// empty data set to reset all DataChanged bits
 _dataChangedNone : AxesGroupStateDataChanged;
  /// internal index for loops
 _idx             : DINT;
END_VAR
// Set internal references 
_stepName      :=   '_stepSyncWorkArea = ';
_rStep       REF=    _stepSyncWorkArea;
_rTimer      REF=   _timerSyncWorkArea;
_rTimeout    REF= _timeoutSyncWorkArea;
_rSyncIdx    REF=     _syncIdxWorkArea;

CASE _rStep
OF    
  0: // Check initialisation configured ?
     // ST-FIX F130: an invalid sync mode (warning of CheckParameterValid) -> no synchronization of the data set
     IF ((( _parCfg.PLC.Parameter.SynchronizationModes.WorkAreas[SyncTime.DURING_START_UP] = SyncMode.NO_SYNCHRONIZATION ) AND
          ( _parCfg.PLC.Parameter.SynchronizationModes.WorkAreas[SyncTime. AFTER_START_UP] = SyncMode.NO_SYNCHRONIZATION )) OR
         ( NOT SyncModesValid( During := _parCfg.PLC.Parameter.SynchronizationModes.WorkAreas[SyncTime.DURING_START_UP],
                               After  := _parCfg.PLC.Parameter.SynchronizationModes.WorkAreas[SyncTime. AFTER_START_UP] ) ))
     THEN
       RETURN;
     END_IF
     
     
     // wait for initialisation done
     IF  ((     AxesGroup.State.RobotData.RCSupportedFunctions. ReadWorkArea ) AND
          (     AxesGroup.State.RobotData.RCSupportedFunctions.WriteWorkArea ) AND
          (     AxesGroup.State.Initialized                                  ) AND 
          ( NOT Error                                                        ))  
     THEN
       // ST-FIX F102: count check after the initialization (HighestXIndex of this connection)
     // Check More Data on RC than on PLC -> Synchronization not possible
     IF (AxesGroup.State.ConfigurationData.HighestWorkAreaIndex > AxesGroup.SystemData.WorkAreasCount)
     THEN
       SetError( ErrorID := RobotLibraryErrorIdEnum.ERR_SYNC_WORKAREA_COUNT_RC_HIGHER_THAN_PLC, Overwrite := FALSE);
       RETURN;
		 END_IF
       // Check PLC WorkAreas < RC WorkAreas and SyncWorkArea enabled ?    
       IF (( AxesGroup.State.DataEnableSync.EnableSyncWorkArea      = TRUE                              )  AND
           ( AxesGroup.Parameter.Rob.Parameter.HighestWorkAreaIndex > AxesGroup.SystemData.WorkAreasMax ))        
       THEN
         SetWarning( WarningID := RobotLibraryWarningIdEnum.WARN_WORK_AREA_ARRAY_TOO_SHORT, Overwrite := TRUE);
       END_IF

       // Create log entry
       CreateLogMessagePara1 ( Timestamp   := SystemTime,
                               MessageType := MessageType.CMD,
                               Severity    := Severity.DEBUG,
                               MessageCode := 0,
                               MessageText := 'SyncWorkArea: Start initial reading of WorkArea from RC',
                               Para1       :=  '');
       
       // init WorkArea number
      _rSyncIdx := DINT_TO_USINT(AxesGroup.SystemData.WorkAreasMin); 
       // init count of unsynchronized elements
       AxesGroup.State.SyncStatePlc.UnSyncNo.WorkArea := 0;
       // set timeout
       SetTimeout(PT := _rTimeout, rTimer := _rTimer);
       // inc step counter
      _rStep := _rStep + 1;
     END_IF     

     
     // Start read WorkArea
  1: IF (( NOT _readWorkArea.Busy  ) AND 
         ( NOT _readWorkArea.Error ) AND
         ( NOT _readWorkArea.Done  ))
     THEN
       // set command parameter
      _readWorkArea.ParCmd.WorkAreaNo := _rSyncIdx;      
       // execute command
      _readWorkArea.Execute := TRUE;
       // set timeout
       SetTimeout(PT := _rTimeout, rTimer := _rTimer);
       // inc step counter
      _rStep := _rStep + 1;
     ELSE
       // check error ? 
       IF ( _readWorkArea.Error ) 
       THEN
         SetWarning ( WarningID := RobotLibraryWarningIdEnum.WARN_WORK_AREA_SYNC_FAILED_BY_ERROR_OF_READ_OR_WRITE_CMD, Overwrite := FALSE );           
       END_IF  
       
       // timeout exceeded ? 
       IF (CheckTimeout(_rTimer) = RobotLibraryConstants.OK)
       THEN
         ErrorID     := RobotLibraryErrorIdEnum.ERR_TIMEOUT_CMD;
         ErrorAddTxt := CONCAT(_stepName, DINT_TO_STRING(_rStep));
       END_IF
     END_IF
 
     
     // Wait WorkArea read
  2: IF (( NOT _readWorkArea.Busy  ) AND
         ( NOT _readWorkArea.Error ) AND
         (     _readWorkArea.Done  ))
     THEN
       // reset execution
      _readWorkArea.Execute := FALSE;
       // set available bit
      _workAreas[_rSyncIdx].Available := TRUE; 
       WorkAreas[_rSyncIdx].Available := TRUE;      
       // Copy data
      _workAreas[_rSyncIdx].Data := _readWorkArea.OutCmd.WorkAreaData;

       // Check WorkArea data is equal ? 
       IF ( NOT IsWorkAreaEqual( Data1 := _workAreas[_rSyncIdx].Data, Data2 := WorkAreas[_rSyncIdx].Data, IgnoreTimestamp := TRUE))
       THEN
         // Reset plc in sync flag
         AxesGroup.State.SyncStatePlc.InSync.WorkArea := FALSE;
         // Set data changed flag
         AxesGroup.State.DataChanged.WorkArea[_rSyncIdx] := TRUE;
         // inc count of unsynchronised plc WorkAreas
         AxesGroup.State.SyncStatePlc.UnSyncNo.WorkArea := AxesGroup.State.SyncStatePlc.UnSyncNo.WorkArea + 1;
        
         // Create log entry
         CreateLogMessagePara1 ( Timestamp   := SystemTime,
                                 MessageType := MessageType.CMD,
                                 Severity    := Severity.DEBUG,
                                 MessageCode := 0,
                                 MessageText := 'SyncWorkArea: Detected a difference in WorkArea[{1}] between PLC and RC',
                                 Para1       :=  DINT_TO_STRING(_rSyncIdx));
        
        
         // Check synchronisation is enabled ? 
         IF ( NOT AxesGroup.State.DataEnableSync.EnableSyncWorkArea )
         THEN
           SetInfo ( InfoID := RobotLibraryInfoIdEnum.INFO_SYNC_WORK_AREA_DISABLED, Overwrite := FALSE );
				 END_IF
         
         // Check user interaction needed ?  
         IF ( AxesGroup.Parameter.PLC.Parameter.SyncUserInteraction.WorkAreas )
         THEN
           SetWarning ( WarningID := RobotLibraryWarningIdEnum.WARN_WORK_AREA_NUMBER_SYNC_ERROR, Overwrite := FALSE );                    
				 END_IF
			 END_IF
             
       // Check all WorkAreas read ? 
       IF ( _rSyncIdx < AxesGroup.State.UnifiedWorkAreaIndex )
       THEN
         // set timeout
         SetTimeout(PT := _rTimeout, rTimer := _rTimer);
         // inc WorkArea index
        _rSyncIdx := _rSyncIdx + 1;
         // dec step counter
        _rStep := _rStep - 1;
       ELSE
         // set timeout
         SetTimeout(PT := _rTimeout, rTimer := _rTimer);
         // inc step counter
        _rStep := _rStep + 1;           
       END_IF
     ELSE
       // check error ? 
       IF (_readWorkArea.Error)
       THEN
         // Set warning
         SetWarning( WarningID := RobotLibraryWarningIdEnum.WARN_WORK_AREA_SYNC_FAILED_BY_ERROR_OF_READ_OR_WRITE_CMD, Overwrite := TRUE);                    
         // reset available bit
         WorkAreas[_rSyncIdx].Available := FALSE;
        _workAreas[_rSyncIdx].Available := FALSE;
       END_IF  
       
       // timeout exceeded ? 
       IF (CheckTimeout(_rTimer) = RobotLibraryConstants.OK)
       THEN
         ErrorID     := RobotLibraryErrorIdEnum.ERR_TIMEOUT_CMD;
         ErrorAddTxt := CONCAT(_stepName, DINT_TO_STRING(_rStep));
       END_IF
     END_IF
     
     
     // Check synchronisation state ? 
  3: IF (( AxesGroup.State.SyncStatePlc.UnSyncNo.WorkArea                                             = 0                           ) OR 
         ( AxesGroup.Parameter.Plc.Parameter.SynchronizationModes.WorkAreas[SyncTime.DURING_START_UP] = SyncMode.NO_SYNCHRONIZATION ))
     THEN
       // Update bit for data in sync
       AxesGroup.State.SyncStatePlc.InSync.WorkArea := (AxesGroup.State.SyncStatePlc.UnSyncNo.WorkArea = 0);
         // ST-FIX F165: synchronization of the start-up phase finished
         AxesGroup.State.Synchronizing.WorkAreas := FALSE;
       // set timeout
       SetTimeout(PT := _rTimeout, rTimer := _rTimer);
       // inc step counter
      _rStep := 10; // -> jump to after startup
            
       // Create log entry
       CreateLogMessagePara1 ( Timestamp   := SystemTime,
                               MessageType := MessageType.CMD,
                               Severity    := Severity.DEBUG,
                               MessageCode := 0,
                               MessageText := 'SyncWorkArea: Synchronization Startup Phase done',
                               Para1       :=  '' );      
     ELSE 
       // Check user interaction needed ? 
       IF ( NOT AxesGroup.Parameter.PLC.Parameter.SyncUserInteraction.WorkAreas )
       THEN
         CASE AxesGroup.Parameter.Plc.Parameter.SynchronizationModes.WorkAreas[SyncTime.DURING_START_UP] OF

           SyncMode.SERVER_TO_CLIENT : 

             // Overwrite PLC data with RC data
             FOR _idx := AxesGroup.SystemData.WorkAreasMin TO MIN(AxesGroup.SystemData.WorkAreasMax, RobotLibraryParameter.WORK_AREAS_MAX - 1) // ST-FIX F18
             DO
               // Overwrite PLC data with RC data
               WorkAreas[_idx] := WorkAreas[_idx];            
						 END_FOR
  
             // Reset data changed flags
             AxesGroup.State.DataChanged.WorkArea := _dataChangedNone.WorkArea;
             // Reset Synchronizing flag
             AxesGroup.State.Synchronizing.WorkAreas := FALSE;
             // Set plc in sync flag
             AxesGroup.State.SyncStatePlc.InSync.WorkArea := TRUE;
             // Reset count of unsynchronised plc WorkAreas
             AxesGroup.State.SyncStatePlc.UnSyncNo.WorkArea := 0;            
             // set timeout
             SetTimeout(PT := _rTimeout, rTimer := _rTimer);
             // inc step counter
            _rStep := 10; // -> jump to after startup         

            // Create log entry
            CreateLogMessagePara3 ( Timestamp   := SystemTime,
                                    MessageType := MessageType.CMD,
                                    Severity    := Severity.DEBUG,
                                    MessageCode := 0,
                                    MessageText := 'SyncWorkArea: Synchronization of WorkAreas triggered by StartUp-Compare, SyncMode = {2}, SyncTime = {3}, SyncDirection = RC -> PLC',
                                    Para1       :=  DINT_TO_STRING(_rSyncIdx),
                                    Para2       :=  SYNC_MODE_TO_STRING(AxesGroup.Parameter.Plc.Parameter.SynchronizationModes.WorkAreas[SyncTime.DURING_START_UP]),
                                    Para3       :=  SYNC_TIME_TO_STRING(SyncTime.DURING_START_UP));
            // Create log entry
            CreateLogMessagePara1 ( Timestamp   := SystemTime,
                                    MessageType := MessageType.CMD,
                                    Severity    := Severity.DEBUG,
                                    MessageCode := 0,
                                    MessageText := 'SyncWorkArea: Applied the initial read WorkArea data from RC',
                                    Para1       :=  '' );

				   SyncMode.CLIENT_TO_SERVER : ;

             // Check conflicts to solve ? 
             FOR _rSyncIdx := 0 TO AxesGroup.State.UnifiedWorkAreaIndex
             DO
               IF ( AxesGroup.State.DataChanged.WorkArea[_rSyncIdx] )
               THEN
                _found := TRUE;
                 EXIT;
		  			   END_IF
             END_FOR
           
             IF ( _found ) 
             THEN
               // Reset plc in sync flag
               AxesGroup.State.SyncStatePlc.InSync.WorkArea := FALSE;
               // Set Synchronizing flag
               AxesGroup.State.Synchronizing.WorkAreas := TRUE;
               // set timeout
               SetTimeout(PT := _rTimeout, rTimer := _rTimer);
               // inc step counter
              _rStep := _rStep +1; // -> write PLC data to RC                  
               // Create log entry
               CreateLogMessagePara3 ( Timestamp   := SystemTime,
                                       MessageType := MessageType.CMD,
                                       Severity    := Severity.DEBUG,
                                       MessageCode := 0,
                                       MessageText := 'SyncWorkArea: Synchronization of WorkArea[{1}] triggered by StartUp-Compare, SyncMode = {2}, SyncTime = {3}, SyncDirection = PLC -> RC',
                                       Para1       :=  DINT_TO_STRING(_rSyncIdx),
                                       Para2       :=  SYNC_MODE_TO_STRING(AxesGroup.Parameter.Plc.Parameter.SynchronizationModes.WorkAreas[SyncTime.DURING_START_UP]),
                                       Para3       :=  SYNC_TIME_TO_STRING(SyncTime.DURING_START_UP));
             ELSE
               // Reset data changed flags
               AxesGroup.State.DataChanged.WorkArea := _dataChangedNone.WorkArea;
               // Reset Synchronizing flag
               AxesGroup.State.Synchronizing.WorkAreas := FALSE;
               // Set plc in sync flag
               AxesGroup.State.SyncStatePlc.InSync.WorkArea := TRUE;
               // Reset count of unsynchronised WorkAreas
               AxesGroup.State.SyncStatePlc.UnSyncNo.WorkArea := 0;
               // set timeout
               SetTimeout(PT := _rTimeout, rTimer := _rTimer);
               // inc step counter
              _rStep := 10; // -> jump to after startup                  
				     END_IF
         ELSE
           // invalid sync mode for startup
           SetWarning( WarningID := RobotLibraryWarningIdEnum.WARN_WORK_AREA_SYNC_MODE_INVALID, Overwrite := TRUE ); // ST-FIX F130: warning instead of the own error
 	       END_CASE
       ELSE
         // ST-FIX F94: the user resolves the conflict with the write / read functions - read the RC data again
         IF ( CheckTimeout(_rTimer) = RobotLibraryConstants.OK )
         THEN
           AxesGroup.State.DataChanged.WorkArea := _dataChangedNone.WorkArea;
           SetTimeout(PT := _rTimeout, rTimer := _rTimer);
          _rStep := 0; // -> read the RC data and compare again
         END_IF
       END_IF
     END_IF  

     
     // Start write WorkArea data  
  4: IF (( NOT _writeWorkArea.Busy  ) AND 
         ( NOT _writeWorkArea.Error ))
     THEN
       // set command parameter
      _writeWorkArea.ParCmd.WorkAreaNo   := _rSyncIdx;      
      _writeWorkArea.ParCmd.WorkAreaData :=  WorkAreas[_rSyncIdx].Data;
       // execute command
      _writeWorkArea.Execute := TRUE;
       // set timeout
       SetTimeout(PT := _rTimeout, rTimer := _rTimer);
       // inc step counter
      _rStep := _rStep + 1;
     ELSE
       // check error ? 
       IF (_writeWorkArea.Error)
       THEN
         ErrorID     := _writeWorkArea.ErrorID;
         ErrorAddTxt := _writeWorkArea.ErrorAddTxt;;
       END_IF  
       
       // timeout exceeded ? 
       IF (CheckTimeout(_rTimer) = RobotLibraryConstants.OK)
       THEN
         ErrorID     := RobotLibraryErrorIdEnum.ERR_TIMEOUT_CMD;
         ErrorAddTxt := CONCAT(_stepName, DINT_TO_STRING(_rStep));
       END_IF
     END_IF
 
     
     // Wait WorkArea data written ?   
  5: IF (( NOT _writeWorkArea.Busy  ) AND
         ( NOT _writeWorkArea.Error ) AND
         (     _writeWorkArea.Done  ))
     THEN
       // execute command
      _writeWorkArea.Execute := FALSE;
       // apply WorkArea data to internal WorkArea data
      _workAreas[_rSyncIdx] := WorkAreas[_rSyncIdx];
       // reset data changed bit 
       AxesGroup.State.DataChanged.WorkArea[_rSyncIdx] := FALSE;
       // dec count of unsynchronised WorkAreas
       AxesGroup.State.SyncStatePlc.UnSyncNo.WorkArea := AxesGroup.State.SyncStatePlc.UnSyncNo.WorkArea - 1;
       // set timeout        
       SetTimeout(PT := _rTimeout, rTimer := _rTimer);
       // dec step counter
      _rStep := _rStep - 2; 
     ELSE
       // check error ? 
       IF (_writeWorkArea.Error)
       THEN
         SetWarning( WarningID := RobotLibraryWarningIdEnum.WARN_WORK_AREA_SYNC_FAILED_BY_ERROR_OF_READ_OR_WRITE_CMD, Overwrite := TRUE);
           // ST-FIX F168: refused by the RC -> warning, go on with the next entry
          _writeWorkArea.Execute := FALSE;
          _workAreas[_rSyncIdx] := WorkAreas[_rSyncIdx];
          AxesGroup.State.DataChanged.WorkArea[_rSyncIdx] := FALSE;
          AxesGroup.State.SyncStatePlc.UnSyncNo.WorkArea := AxesGroup.State.SyncStatePlc.UnSyncNo.WorkArea - 1;
           SetTimeout(PT := _rTimeout, rTimer := _rTimer);
          _rStep := _rStep - 2;           
       END_IF  
       
       // timeout exceeded ? 
       IF (CheckTimeout(_rTimer) = RobotLibraryConstants.OK)
       THEN
         ErrorID     := RobotLibraryErrorIdEnum.ERR_TIMEOUT_CMD;
         ErrorAddTxt := CONCAT(_stepName, DINT_TO_STRING(_rStep));
       END_IF
     END_IF

     
  // --------------------------------------------
  // SyncMode after startup : 
  // --------------------------------------------
         
  10 : // check synchronisation active ? 
       // ST-FIX F93: compare also with NO_SYNCHRONIZATION (no transfer, see the CASE below)
       
       // reset count of unsynchronised WorkAreas
       AxesGroup.State.SyncStatePlc.UnSyncNo.WorkArea := 0;

       // Check all WorkArea datas
       FOR _rSyncIdx := 0 TO AxesGroup.State.UnifiedWorkAreaIndex
       DO
         // compare WorkArea data
         AxesGroup.State.DataChanged.WorkArea[_rSyncIdx] := NOT IsWorkAreaEqual( Data1 := WorkAreas[_rSyncIdx].Data, Data2 := _workAreas[_rSyncIdx].Data, IgnoreTimestamp := TRUE (* ST-FIX F57 *));

         // Check WorkArea data changed ? 
         IF (AxesGroup.State.DataChanged.WorkArea[_rSyncIdx])
         THEN
           // inc count of unsynchronised plc WorkAreas
           AxesGroup.State.SyncStatePlc.UnSyncNo.WorkArea := AxesGroup.State.SyncStatePlc.UnSyncNo.WorkArea + 1;
           // Create log entry
           CreateLogMessagePara2 ( Timestamp   := SystemTime,
                                   MessageType := MessageType.CMD,
                                   Severity    := Severity.DEBUG,
                                   MessageCode := 0,
                                   MessageText := 'SyncWorkArea: Detected a local change of WorkArea[{1}] on PLC, SyncTime = {2}',
                                   Para1       :=  DINT_TO_STRING(_rSyncIdx),    
                                   Para2       :=  SYNC_TIME_TO_STRING(SyncTime.AFTER_START_UP));       
				 END_IF

         // Update plc in sync flag
         AxesGroup.State.SyncStatePlc.InSync.WorkArea := (AxesGroup.State.SyncStatePlc.UnSyncNo.WorkArea = 0); 
	     END_FOR

       // Check synchronization is needed ? 
       IF ( NOT AxesGroup.State.SyncStatePlc.InSync.WorkArea ) XOR  
          ( NOT AxesGroup.State.SyncStateRc .InSync.WorkArea )
       THEN
         CASE AxesGroup.Parameter.Plc.Parameter.SynchronizationModes.WorkAreas[SyncTime.AFTER_START_UP] 
         OF         
           // NO_SYNCHRONIZATION
           SyncMode.NO_SYNCHRONIZATION : ; // no further action 
           
           // CLIENT_TO_SERVER
           SyncMode.CLIENT_TO_SERVER :
             // set timeout
             SetTimeout(PT := _rTimeout, rTimer := _rTimer);
             // inc step counter
            _rStep := 11;
  
           // SERVER_TO_CLIENT
           SyncMode.SERVER_TO_CLIENT :
             // set timeout
             SetTimeout(PT := _rTimeout, rTimer := _rTimer);
             // inc step counter
            _rStep := 12;
  
           // AUTOMATIC
           SyncMode.AUTOMATIC : 
             // set timeout
             SetTimeout(PT := _rTimeout, rTimer := _rTimer);
             // inc step counter
            _rStep := 13;
         END_CASE
       ELSE
         // datas changeḍ on both sides ? -> Warning 
         IF (( NOT AxesGroup.State.SyncStatePlc.InSync.WorkArea ) AND  
             ( NOT AxesGroup.State.SyncStateRc .InSync.WorkArea ))
         THEN
           // ST-FIX F58: CLIENT_TO_SERVER / SERVER_TO_CLIENT decide the direction also if both sides changed
CASE AxesGroup.Parameter.Plc.Parameter.SynchronizationModes.WorkAreas[SyncTime.AFTER_START_UP] OF
  SyncMode.CLIENT_TO_SERVER : _rStep := 11;
  SyncMode.SERVER_TO_CLIENT : _rStep := 12;
ELSE
  SetWarning( WarningID := RobotLibraryWarningIdEnum.WARN_WORK_AREA_SYNC_BOTH_SIDES_CHANGED, Overwrite := TRUE);
END_CASE
         END_IF
       END_IF


  // ------------------------------------------
  // SyncMode : CLIENT_TO_SERVER 
  // ------------------------------------------  
  11 : // Conflict triggerd by PLC ?  
       IF ( NOT AxesGroup.State.SyncStatePlc.InSync.WorkArea )
       THEN
         // search for changed index  
         FOR _rSyncIdx := 0 TO AxesGroup.State.UnifiedWorkAreaIndex
         DO
           IF ( AxesGroup.State.DataChanged.WorkArea[_rSyncIdx] )
           THEN
             // set timeout
             SetTimeout(PT := _rTimeout, rTimer := _rTimer);
             // inc step counter
            _rStep := 30; // -> write PLC data to RC                  
             EXIT;             
					 END_IF
         END_FOR
         
         // Create log entry
         CreateLogMessagePara3 ( Timestamp   := SystemTime,
                                 MessageType := MessageType.CMD,
                                 Severity    := Severity.DEBUG,
                                 MessageCode := 0,
                                 MessageText := 'SyncWorkArea: Synchronization of WorkArea[{1}] triggered by PLC, SyncMode = {2}, SyncTime = {3}, SyncDirection = PLC -> RC',
                                 Para1       :=  DINT_TO_STRING(_rSyncIdx),
                                 Para2       :=  SYNC_MODE_TO_STRING(AxesGroup.Parameter.Plc.Parameter.SynchronizationModes.WorkAreas[SyncTime.AFTER_START_UP]),
                                 Para3       :=  SYNC_TIME_TO_STRING(SyncTime.AFTER_START_UP));
                                 RETURN;
       END_IF
   
       // Conflict triggered by RC ?
       IF ( NOT AxesGroup.State.SyncStateRc.InSync.WorkArea )
       THEN
         // get changed index 
        _rSyncIdx :=  LIMIT(0, AxesGroup.State.SyncStateRc.UnSyncNo.WorkArea, AxesGroup.State.UnifiedWorkAreaIndex);
         // set timeout
         SetTimeout(PT := _rTimeout, rTimer := _rTimer);
         // inc step counter
        _rStep := 30; // -> write PLC data to RC

         // Create log entry
         CreateLogMessagePara3 ( Timestamp   := SystemTime,
                                 MessageType := MessageType.CMD,
                                 Severity    := Severity.DEBUG,
                                 MessageCode := 0,
                                 MessageText := 'SyncWorkArea: Synchronization of WorkArea[{1}] triggered by RC, SyncMode = {2}, SyncTime = {3}, SyncDirection = PLC -> RC',
                                 Para1       :=  DINT_TO_STRING(_rSyncIdx),
                                 Para2       :=  SYNC_MODE_TO_STRING(AxesGroup.Parameter.Plc.Parameter.SynchronizationModes.WorkAreas[SyncTime.AFTER_START_UP]),
                                 Para3       :=  SYNC_TIME_TO_STRING(SyncTime.AFTER_START_UP));
                                 RETURN;
			 END_IF
       
       // set timeout
       SetTimeout(PT := _rTimeout, rTimer := _rTimer);
       // jump back
      _rStep := 10;

       
  // ------------------------------------------
  // SyncMode : SERVER_TO_CLIENT 
  // ------------------------------------------
  12 : // Conflict triggerd by PLC ?  
       IF ( NOT AxesGroup.State.SyncStatePlc.InSync.WorkArea )
       THEN
         // search for changed index  
         FOR _rSyncIdx := 0 TO AxesGroup.State.UnifiedWorkAreaIndex
         DO
           IF ( AxesGroup.State.DataChanged.WorkArea[_rSyncIdx] )
           THEN
             // set timeout
             SetTimeout(PT := _rTimeout, rTimer := _rTimer);
             // inc step counter
            _rStep := 20; // -> read RC data and write it to PLC                  
             EXIT;
					 END_IF
         END_FOR

         // Create log entry
         CreateLogMessagePara3 ( Timestamp   := SystemTime,
                                 MessageType := MessageType.CMD,
                                 Severity    := Severity.DEBUG,
                                 MessageCode := 0,
                                 MessageText := 'SyncWorkArea: Synchronization of WorkArea[{1}] triggered by PLC, SyncMode = {2}, SyncTime = {3}, SyncDirection = RC -> PLC',
                                 Para1       :=  DINT_TO_STRING(_rSyncIdx),
                                 Para2       :=  SYNC_MODE_TO_STRING(AxesGroup.Parameter.Plc.Parameter.SynchronizationModes.WorkAreas[SyncTime.AFTER_START_UP]),
                                 Para3       :=  SYNC_TIME_TO_STRING(SyncTime.AFTER_START_UP));
                                 RETURN;
       END_IF
   
       // Conflict triggered by RC ?
       IF ( NOT AxesGroup.State.SyncStateRc.InSync.WorkArea )
       THEN
         // get changed index 
        _rSyncIdx := LIMIT(0, AxesGroup.State.SyncStateRc.UnSyncNo.WorkArea, AxesGroup.State.UnifiedWorkAreaIndex);
         // set timeout
         SetTimeout(PT := _rTimeout, rTimer := _rTimer);
         // inc step counter
        _rStep := 20; // -> read RC data and write it to PLC

         // Create log entry
         CreateLogMessagePara3 ( Timestamp   := SystemTime,
                                 MessageType := MessageType.CMD,
                                 Severity    := Severity.DEBUG,
                                 MessageCode := 0,
                                 MessageText := 'SyncWorkArea: Synchronization of WorkArea[{1}] triggered by RC, SyncMode = {2}, SyncTime = {3}, SyncDirection = RC -> PLC',
                                 Para1       :=  DINT_TO_STRING(_rSyncIdx),
                                 Para2       :=  SYNC_MODE_TO_STRING(AxesGroup.Parameter.Plc.Parameter.SynchronizationModes.WorkAreas[SyncTime.AFTER_START_UP]),
                                 Para3       :=  SYNC_TIME_TO_STRING(SyncTime.AFTER_START_UP));
                                 RETURN;
			 END_IF
       
       // set timeout
       SetTimeout(PT := _rTimeout, rTimer := _rTimer);
       // jump back
      _rStep := 10;
  

  // ------------------------------------------
  // SyncMode : AUTOMATIC 
  // ------------------------------------------
  13 : // Conflict triggerd by PLC ?  
       IF ( NOT AxesGroup.State.SyncStatePlc.InSync.WorkArea )
       THEN
         // search for changed index  
         FOR _rSyncIdx := 0 TO AxesGroup.State.UnifiedWorkAreaIndex
         DO
           IF ( AxesGroup.State.DataChanged.WorkArea[_rSyncIdx] )
           THEN
             // set timeout
             SetTimeout(PT := _rTimeout, rTimer := _rTimer);
             // inc step counter
            _rStep := 30; // -> write PLC data to RC                  
             EXIT;
					 END_IF
         END_FOR
         
         // Create log entry
         CreateLogMessagePara3 ( Timestamp   := SystemTime,
                                 MessageType := MessageType.CMD,
                                 Severity    := Severity.DEBUG,
                                 MessageCode := 0,
                                 MessageText := 'SyncWorkArea: Synchronization of WorkArea[{1}] triggered by PLC, SyncMode = {2}, SyncTime = {3}, SyncDirection = PLC -> RC',
                                 Para1       :=  DINT_TO_STRING(_rSyncIdx),
                                 Para2       :=  SYNC_MODE_TO_STRING(AxesGroup.Parameter.Plc.Parameter.SynchronizationModes.WorkAreas[SyncTime.AFTER_START_UP]),
                                 Para3       :=  SYNC_TIME_TO_STRING(SyncTime.AFTER_START_UP));
                                 RETURN;
       END_IF
   
       // Conflict triggered by RC ?
       IF ( NOT AxesGroup.State.SyncStateRc.InSync.WorkArea )
       THEN
         // get changed index 
        _rSyncIdx := LIMIT(0, AxesGroup.State.SyncStateRc.UnSyncNo.WorkArea, AxesGroup.State.UnifiedWorkAreaIndex);
         // set timeout
         SetTimeout(PT := _rTimeout, rTimer := _rTimer);
         // inc step counter
        _rStep := 20; // -> read RC data an write it to PLC

         // Create log entry
         CreateLogMessagePara3 ( Timestamp   := SystemTime,
                                 MessageType := MessageType.CMD,
                                 Severity    := Severity.DEBUG,
                                 MessageCode := 0,
                                 MessageText := 'SyncWorkArea: Synchronization of WorkArea[{1}] triggered by RC, SyncMode = {2}, SyncTime = {3}, SyncDirection = RC -> PLC',
                                 Para1       :=  DINT_TO_STRING(_rSyncIdx),
                                 Para2       :=  SYNC_MODE_TO_STRING(AxesGroup.Parameter.Plc.Parameter.SynchronizationModes.WorkAreas[SyncTime.AFTER_START_UP]),
                                 Para3       :=  SYNC_TIME_TO_STRING(SyncTime.AFTER_START_UP));
                                 RETURN;
			 END_IF
       
       // set timeout
       SetTimeout(PT := _rTimeout, rTimer := _rTimer);
       // jump back
      _rStep := 10; // ST-FIX F95: was commented out


  // ------------------------------------------
  // Read Data from RC and write it to PLC
  // ------------------------------------------
  20 : IF (( NOT _readWorkArea.Busy  ) AND 
           ( NOT _readWorkArea.Error ))
       THEN
         // set command parameter
        _readWorkArea.ParCmd.WorkAreaNo := _rSyncIdx;      
         // execute command
        _readWorkArea.Execute := TRUE;
         // set timeout
         SetTimeout(PT := _rTimeout, rTimer := _rTimer);
         // inc step counter
        _rStep := _rStep + 1;
       ELSE
         // check error ? 
         IF (_readWorkArea.Error)
         THEN
           ErrorID     := _readWorkArea.ErrorID;
           ErrorAddTxt := _readWorkArea.ErrorAddTxt;
         END_IF  
       
         // timeout exceeded ? 
         IF (CheckTimeout(_rTimer) = RobotLibraryConstants.OK)
         THEN
           ErrorID     := RobotLibraryErrorIdEnum.ERR_TIMEOUT_CMD;
           ErrorAddTxt := CONCAT(_stepName, DINT_TO_STRING(_rStep));
         END_IF
       END_IF
 
  21 : IF (( NOT _readWorkArea.Busy  ) AND
           ( NOT _readWorkArea.Error ) AND
           (     _readWorkArea.Done  ))
       THEN
         // reset execution
        _readWorkArea.Execute := FALSE;
         // ST-FIX F107: AUTOMATIC - the PLC data were changed while the RC data were read: the PLC
         // change is the most recent one and is written to the RC instead of being overwritten
         IF ( AxesGroup.Parameter.Plc.Parameter.SynchronizationModes.WorkAreas[SyncTime.AFTER_START_UP] = SyncMode.AUTOMATIC ) AND
            ( NOT IsWorkAreaEqual( Data1 := WorkAreas[_rSyncIdx].Data, Data2 := _workAreas[_rSyncIdx].Data, IgnoreTimestamp := TRUE ))
         THEN
           // set timeout
           SetTimeout(PT := _rTimeout, rTimer := _rTimer);
           // -> write PLC data to RC
          _rStep := 30;
           RETURN;
         END_IF
         // update internal WorkArea data
         WorkAreas[_rSyncIdx].Data := _readWorkArea.OutCmd.WorkAreaData;         
        _workAreas[_rSyncIdx].Data := _readWorkArea.OutCmd.WorkAreaData;
         // set available bit
         WorkAreas[_rSyncIdx].Available := TRUE;
        _workAreas[_rSyncIdx].Available := TRUE;
         // set timeout
         SetTimeout(PT := _rTimeout, rTimer := _rTimer);
         // inc step counter
        // ST-FIX F20: write the RC data back to reset DataChanged on the RC (spec 5.6.7.4.2)
        IF ( AxesGroup.State.RobotData.RCSupportedFunctions.WriteWorkArea )
        THEN
          _rStep := 30;
        ELSE
          _rStep := 10;
        END_IF // -> jump to after startup           
       ELSE
         // check error ? 
         IF (_readWorkArea.Error)
         THEN
           ErrorID     := _readWorkArea.ErrorID;
           ErrorAddTxt := _readWorkArea.ErrorAddTxt;           
           // reset available bit
           WorkAreas[_rSyncIdx].Available := FALSE;
          _workAreas[_rSyncIdx].Available := FALSE;
         END_IF  
       
         // timeout exceeded ? 
         IF (CheckTimeout(_rTimer) = RobotLibraryConstants.OK)
         THEN
           ErrorID     := RobotLibraryErrorIdEnum.ERR_TIMEOUT_CMD;
           ErrorAddTxt := CONCAT(_stepName, DINT_TO_STRING(_rStep));
         END_IF
       END_IF


  // ------------------------------------------
  // Write data from PLC to RC
  // ------------------------------------------
  30 : IF (( NOT _writeWorkArea.Busy  ) AND 
           ( NOT _writeWorkArea.Error ))
       THEN
         // set command parameter
        _writeWorkArea.ParCmd.WorkAreaNo   := _rSyncIdx;      
        _writeWorkArea.ParCmd.WorkAreaData :=  WorkAreas[_rSyncIdx].Data;
         // execute command
        _writeWorkArea.Execute := TRUE;
         // set timeout
         SetTimeout(PT := _rTimeout, rTimer := _rTimer);
         // inc step counter
        _rStep := _rStep + 1;
       ELSE
         // check error ? 
         IF (_writeWorkArea.Error)
         THEN
           ErrorID     := _writeWorkArea.ErrorID;
           ErrorAddTxt := _writeWorkArea.ErrorAddTxt;;
         END_IF  
       
         // timeout exceeded ? 
         IF (CheckTimeout(_rTimer) = RobotLibraryConstants.OK)
         THEN
           ErrorID     := RobotLibraryErrorIdEnum.ERR_TIMEOUT_CMD;
           ErrorAddTxt := CONCAT(_stepName, DINT_TO_STRING(_rStep));
         END_IF
       END_IF
 
  31 : IF (( NOT _writeWorkArea.Busy  ) AND
           ( NOT _writeWorkArea.Error ) AND
           (     _writeWorkArea.Done  ))
       THEN
         // execute command
        _writeWorkArea.Execute := FALSE;      
         // update internal WorkArea data
        _workAreas[_rSyncIdx] := WorkAreas[_rSyncIdx]; 
         // set available bit
         WorkAreas[_rSyncIdx].Available := TRUE; 
        _workAreas[_rSyncIdx].Available := TRUE;         
         // set timeout
         SetTimeout(PT := _rTimeout, rTimer := _rTimer);
         // inc step counter
        _rStep := 10; // -> jump to after startup;           
       ELSE
         // check error ? 
         IF (_writeWorkArea.Error)
         THEN
           SetWarning( WarningID := RobotLibraryWarningIdEnum.WARN_WORK_AREA_SYNC_FAILED_BY_ERROR_OF_READ_OR_WRITE_CMD, Overwrite :=  TRUE);    
           // reset available bit
           WorkAreas[_rSyncIdx].Available := FALSE;
          _workAreas[_rSyncIdx].Available := FALSE;
         END_IF  
       
         // timeout exceeded ? 
         IF (CheckTimeout(_rTimer) = RobotLibraryConstants.OK)
         THEN
           ErrorID     := RobotLibraryErrorIdEnum.ERR_TIMEOUT_CMD;
           ErrorAddTxt := CONCAT(_stepName, DINT_TO_STRING(_rStep));
         END_IF
       END_IF
       
ELSE
  // invalid step
  ErrorID     := RobotLibraryErrorIdEnum.ERR_INVALID_STEP;
  ErrorAddTxt := CONCAT(_stepName , DINT_TO_STRING(_stepCmd));
END_CASE
END_METHOD

METHOD PRIVATE HandleTelegramStateCtrl
VAR_INPUT
END_VAR
// Telegram Control
// ----------------
IF ( _lastTelegramControl <> GetHalfeByteLo(Telegram.PlcToRob.Header.AxesGroupID_Control))
THEN
  // Create log entry
  CreateLogMessagePara2 ( Timestamp   := SystemTime,
                          MessageType := MessageType.CMD,
                          Severity    := Severity.INFO,
                          MessageCode := 0,
                          MessageText := 'SRCI Interface control changed from {1} to {2}',
                          Para1       := TELEGRAM_CONTROL_TO_STRING(_lastTelegramControl),
                          Para2       := TELEGRAM_CONTROL_TO_STRING(GetHalfeByteLo(Telegram.PlcToRob.Header.AxesGroupID_Control)));

  _lastTelegramControl := GetHalfeByteLo(Telegram.PlcToRob.Header.AxesGroupID_Control);
END_IF


// Telegram State
// ----------------
IF ( _lastTelegramState <> Telegram.RobToPlc.Header.TelegramState)
THEN
  // Create log entry
  CreateLogMessagePara2 ( Timestamp   := SystemTime,
                          MessageType := MessageType.CMD,
                          Severity    := Severity.INFO,
                          MessageCode := 0,
                          MessageText := 'SRCI Interface state changed from {1} to {2}',
                          Para1       := TELEGRAM_STATE_TO_STRING(_lastTelegramState),
                          Para2       := TELEGRAM_STATE_TO_STRING(Telegram.RobToPlc.Header.TelegramState));


  // Check Interface changed after being initialized ?  
  IF ((  Enable                                                                          ) AND
      ( _lastTelegramState                      = TelegramState.INITIALIZED              ) AND  
     ((  Telegram.RobToPlc.Header.TelegramState = TelegramState.READY_FOR_INITIALIZATION ) OR
      (  Telegram.RobToPlc.Header.TelegramState = TelegramState.READY_TO_RESUME          )))
  THEN
    // the error 16#80A7 (interface reset after the initialization) is set in OnCall (ST-FIX F65)
    ;
	END_IF

  // apply new telegram state
 _lastTelegramState := Telegram.RobToPlc.Header.TelegramState;
END_IF
END_METHOD

METHOD HandleUserData
VAR_IN_OUT
   /// Robot assignment of function
  AxesGroup    : AxesGroup;
  ///  User data stored on the PLC according to Table 6-10
  UserData     : UserData;
END_VAR
// Common
UserData.LogLevel                          := LogLevel;

UserData.PLCManufacturedID                 := _parCfg.Plc.Parameter.ManufacturedID;
UserData.PLCOrderID                        := _parCfg.Plc.Parameter.OrderID;
UserData.PLCSerialNumber                   := _parCfg.Plc.Parameter.SerialNumber;
UserData.PLCFirmwareVersion                := _parCfg.Plc.Parameter.FirmwareVersion;
UserData.PLCInterfaceVersion               := _parCfg.Plc.Parameter.InterfaceVersion;
UserData.PLCLibraryVersion                 :=  RobotLibraryConstants.PLCLibraryVersion;
                                           
// Communication                           
UserData.LifeSignTimeOut                   := _parCfg.Com.LifeSignTimeOut;
                                           
// Plc Parameter                           
UserData.SynchronizationModes              := _parCfg.Plc.Parameter.SynchronizationModes;
UserData.EnableSync                        :=  SyncModesToDataEnableSync(Value := _parCfg.Plc.Parameter.SynchronizationModes);
                                           
// Robot Parameter                         
UserData.DelayTime                         := _parCfg.Rob.Parameter.DelayTime;
UserData.WaitForNrOfCmd                    := _parCfg.Rob.Parameter.WaitForNrOfCmd;
UserData.WaitAtBlendingZone                := _parCfg.Rob.Parameter.WaitAtBlendingZone;
UserData.AllowSecSeqWhileSubprogram        := _parCfg.Rob.Parameter.AllowSecSeqWhileSubprogram;
UserData.AllowDynamicBlending              := _parCfg.Rob.Parameter.AllowDynamicBlending;
UserData.SyncReaction                      := _parCfg.Rob.Parameter.SyncReaction;
UserData.SyncDelay                         := _parCfg.Rob.Parameter.SyncDelay;
UserData.MessageLevel                      := _parcfg.Rob.Parameter.MessageLevel;

// ReadRobotData
UserData.RCManufacturer                    := AxesGroup.State.RobotData.RCManufacturer; 
UserData.RCOrderID                         := AxesGroup.State.RobotData.RCOrderID; 
UserData.RCSerialNumber                    := AxesGroup.State.RobotData.RCSerialNumber;
UserData.RASerialNumber                    := AxesGroup.State.RobotData.RASerialNumber;
UserData.RCFirmwareVersion                 := AxesGroup.State.RobotData.RCFirmwareVersion;

UserData.RCInterpreterVersion := AxesGroup.State.RobotData.RCInterpreterVersionNumber; // ST-FIX F163: was characters 1/2/3 of the text

UserData.AxisJointUsed                     := AxesGroup.State.RobotData.AxisJointUsed;
UserData.AxisExternalUsed                  := AxesGroup.State.RobotData.AxisExternalUsed;
UserData.AxisJointUnit                     := AxesGroup.State.RobotData.AxisJointUnit;
UserData.AxisExternalUnit                  := AxesGroup.State.RobotData.AxisExternalUnit;
UserData.RCSupportedFunctions              := AxesGroup.State.RobotData.RCSupportedFunctions;
                                           
UserData.BrakeTestRequired                 := AxesGroup.State.ConfigurationData.BrakeTestRequired;
UserData.PathAccuracyMode                  := AxesGroup.State.ConfigurationData.PathAccuracyMode;
UserData.AvoidSingularity                  := AxesGroup.State.ConfigurationData.AvoidSingularity;
UserData.ConstantVelocitySupported         := AxesGroup.State.ConfigurationData.ConstantVelocitySupported;
UserData.StepModeExactStopActive           := AxesGroup.State.ConfigurationData.StepModeExactStopActive;
UserData.StepModeBlendingActive            := AxesGroup.State.ConfigurationData.StepModeBlendingActive;
UserData.AcceleratingSupported             := AxesGroup.State.ConfigurationData.AcceleratingSupported;
UserData.DeceleratingSupported             := AxesGroup.State.ConfigurationData.DecceleratingSupported;
                                           
UserData.Initialized                       := Initialized;
UserData.Synchronized                      := Synchronized;
                                           
// Cyclic data                             
UserData.RCSRCIVersion                     := AxesGroup.Cyclic.RobToPlc.SRCIVersion;
UserData.IsMoving                          := AxesGroup.Cyclic.RobToPlc.StatusRobotArm.IsMoving;
UserData.PrimarySequencePaused             := AxesGroup.Cyclic.RobToPlc.StatusRobotArm.PrimarySequencePaused;
UserData.InPrimaryPos                      := AxesGroup.Cyclic.RobToPlc.StatusRobotArm.InPrimaryPos;
UserData.SecondarySequenceActive           := AxesGroup.Cyclic.RobToPlc.StatusRobotArm.SecondarySequenceActive;
UserData.ErrorPending                      := AxesGroup.Cyclic.RobToPlc.StatusRobotArm.ErrorPending;
UserData.RestartInProgress                 := AxesGroup.Cyclic.RobToPlc.StatusRobotArm.RestartInProgress;
UserData.Enabled                           := AxesGroup.Cyclic.RobToPlc.StatusRobotArm.Enabled;
UserData.Idle                              := AxesGroup.Cyclic.RobToPlc.StatusRobotArm.RaSequenceState = RaSequenceState.IDLE;
UserData.Executing                         := AxesGroup.Cyclic.RobToPlc.StatusRobotArm.RaSequenceState = RaSequenceState.EXECUTING;
UserData.Interrupted                       := AxesGroup.Cyclic.RobToPlc.StatusRobotArm.RaSequenceState = RaSequenceState.INTERRUPTED;
UserData.IsBlending                        := AxesGroup.Cyclic.RobToPlc.StatusRobotArm.IsBlending;  
UserData.OperationMode                     := AxesGroup.Cyclic.RobToPlc.StatusRobotArm.OperationMode;
UserData.CollisionDetectionEnabled         := AxesGroup.Parameter.Rob.Parameter.CollisionDetectionEnabled; // ST-FIX F169: the status word bit is always FALSE
UserData.CollisionDetected                 := AxesGroup.Cyclic.RobToPlc.StatusRobotArm.CollisionDetected;
UserData.RestartRequested                  := AxesGroup.Cyclic.RobToPlc.StatusRobotArm.RestartRequested;
UserData.Accelerating                      := AxesGroup.Cyclic.RobToPlc.StatusRobotArm.Accelerating;
UserData.Decelerating                      := AxesGroup.Cyclic.RobToPlc.StatusRobotArm.Decelerating;
UserData.ConstantVelocity                  := AxesGroup.Cyclic.RobToPlc.StatusRobotArm.ConstantVelocity;
UserData.ActualOverride                    := PERCENT_UINT_TO_REAL( Value := AxesGroup.Cyclic.RobToPlc.Override, IsOptional := FALSE);

// Cyclic optional data
UserData.CartesianPosition                 := AxesGroup.CyclicOptional.RobToPlc.CartesianPosition;
UserData.ExtCartesianPosition              := AxesGroup.CyclicOptional.RobToPlc.CartesianPositionExt;  
UserData.JointPosition                     := AxesGroup.CyclicOptional.RobToPlc.JointPosition;
UserData.ExtJointPosition                  := AxesGroup.CyclicOptional.RobToPlc.JointPositionExt;

// Synchronizing
UserData.ToolDataSynchronizing             := AxesGroup.State.Synchronizing.Tool;
UserData.FrameDataSynchronizing            := AxesGroup.State.Synchronizing.Frame;
UserData.LoadDataSynchronizing             := AxesGroup.State.Synchronizing.Load;
UserData.WorkAreaDataSynchronizing         := AxesGroup.State.Synchronizing.WorkAreas;
UserData.SWLimitsSynchronizing             := AxesGroup.State.Synchronizing.SwLimits;
UserData.DefaultDynamicsSynchronizing      := AxesGroup.State.Synchronizing.DefaultDynamics;
UserData.ReferenceDynamicsSynchronizing    := AxesGroup.State.Synchronizing.ReferenceDynamics;


UserData.ActivateTwoSequences              := _parCfg.Com.TwoSequences;
UserData.ReadingCartesianPosition          :=  AxesGroup.State.ReadingCartesianPosition;
UserData.ReadingExtCartesianPosition       :=  AxesGroup.State.ReadingCartesianPositionExt;
UserData.ReadingJointPosition              :=  AxesGroup.State.ReadingJointPosition;
UserData.ReadingExtJointPosition           :=  AxesGroup.State.ReadingJointPositionExt;
END_METHOD

PROPERTY PROTECTED HasError : Bool
GET
HasError := ErrorID <> RobotLibraryErrorIdEnum.NO_ERROR;
END_GET
END_PROPERTY

PROPERTY PROTECTED HasInfo : BOOL
GET
HasInfo := InfoID <> RobotLibraryInfoIdEnum.NO_INFO;
END_GET
END_PROPERTY

PROPERTY PROTECTED HasWarning : BOOL
GET
HasWarning := WarningID <> RobotLibraryWarningIdEnum.NO_WARNING;
END_GET
END_PROPERTY

METHOD PRIVATE OnCall
VAR_IN_OUT
   /// Robot assignment of function
  AxesGroup : AxesGroup;
END_VAR
// map numeric value to enum, so that the corresponding message text is directly shown by the tooltip
ErrorIdEnum   := ErrorId;
WarningIdEnum := WarningId;
InfoIdEnum    := InfoId;

Error := HasError;

// Check Payload and In/Out data size
IF (( ROBOT_IN_DATA_SIZE  < 64 ) OR
    ( ROBOT_OUT_DATA_SIZE < 64 ))
THEN
  SetError(ErrorID := RobotLibraryErrorIdEnum.ERR_INVALID_LIBRARY_PARA, Overwrite := TRUE );
  RETURN;
END_IF


// Check AxesGroupID valid
IF (( AxesGroupID < RobotLibraryConstants.AXES_GROUP_ID_MIN ) OR
    ( AxesGroupID > RobotLibraryConstants.AXES_GROUP_ID_MAX ))
THEN
  // ST-FIX F138: client error of the specification (16#80AA, table 7-2) instead of the internal ID 3
  SetError( ErrorID := RobotLibraryErrorIdEnum.ERR_AXESGROUP_ID_INVALID_0x80AA, Overwrite := TRUE );
  RETURN;
END_IF


// Reset flag for initialization / Synchronization
IF ( Initialized OR Synchronized) AND ( AxesGroup.Cyclic.RobToPlc.TelegramState <> TelegramState.INITIALIZED)
THEN
  // Reset initialized flag
  Initialized := FALSE;
  // Reset Synchronized flag
  Synchronized := FALSE;
  // Set error 
  // ST-FIX F65: reason of the loss of the initialization (table 7-2): RI error of the RC in the
  // telegram state (16#A1..16#AD), interface reset by the RC (16#80A7) or unknown (16#80A2)
  IF (( AxesGroup.Cyclic.RobToPlc.TelegramState >= TelegramState.ERROR_161_TELEGRAM_CONTROL_MISMATCH_TELEGRAM_STATE ) AND
      ( AxesGroup.Cyclic.RobToPlc.TelegramState <= TelegramState.ERROR_173_SERVER_CONNECTION_LOST                   ))
  THEN
    SetError( ErrorID := AxesGroup.Cyclic.RobToPlc.TelegramState, Overwrite := TRUE );
    // Create log entry
    CreateLogMessagePara1 ( Timestamp   := SystemTime,
                            MessageType := MessageType.CMD,
                            Severity    := Severity.ERROR,
                            MessageCode := ErrorID,
                            MessageText := 'Initialization lost: RI error {1} of the RC',
                            Para1       := TELEGRAM_STATE_TO_STRING(AxesGroup.Cyclic.RobToPlc.TelegramState));
  ELSIF (( AxesGroup.Cyclic.RobToPlc.TelegramState = TelegramState.READY_FOR_INITIALIZATION ) OR
         ( AxesGroup.Cyclic.RobToPlc.TelegramState = TelegramState.READY_TO_RESUME          ))
  THEN
    SetError( ErrorID := RobotLibraryErrorIdEnum.ERR_INTERFACE_WAS_RESET_AFTER_INIT_0x80A7, Overwrite := TRUE );
    // Create log entry
    CreateLogMessagePara1 ( Timestamp   := SystemTime,
                            MessageType := MessageType.CMD,
                            Severity    := Severity.ERROR,
                            MessageCode := ErrorID,
                            MessageText := 'Initialization lost: interface was reset by the RC (state {1})',
                            Para1       := TELEGRAM_STATE_TO_STRING(AxesGroup.Cyclic.RobToPlc.TelegramState));
  ELSE
    SetError( ErrorID := RobotLibraryErrorIdEnum.ERR_INIT_LOST_UNKNOWN_0x80A2, Overwrite := TRUE );
    // Create log entry
    CreateLogMessagePara1 ( Timestamp   := SystemTime,
                            MessageType := MessageType.CMD,
                            Severity    := Severity.ERROR,
                            MessageCode := ErrorID,
                            MessageText := 'Initialization lost: unknown reason (state {1})',
                            Para1       := TELEGRAM_STATE_TO_STRING(AxesGroup.Cyclic.RobToPlc.TelegramState));
  END_IF
END_IF


// Warning for ACR Registers running low
IF ( AxesGroup.Acyclic.ActiveCommandRegister.CurrentAcrUsagePercent > RobotLibraryParameter.ACR_USAGE_WARNING_LIMIT )
THEN
  SetWarning( WarningID := RobotLibraryWarningIdEnum.WARN_ACR_FREE_ENTRIES_LOW, Overwrite := TRUE);  
END_IF

// Check ToolData boundary
IF ( AxesGroup.SystemData.ToolDataMin  <> 0 )  
THEN
  SetWarning( WarningID := RobotLibraryWarningIdEnum.WARN_TOOL_DATA_ARRAY_NOT_START_AT_ZERO, Overwrite := FALSE );
END_IF

// Check FrameData boundary
IF ( AxesGroup.SystemData.FrameDataMin <> 0 ) AND ( NOT HasWarning )  
THEN
  SetWarning( WarningID := RobotLibraryWarningIdEnum.WARN_FRAME_DATA_ARRAY_NOT_START_AT_ZERO, Overwrite := FALSE );
END_IF

// Check WorkAreas boundary
IF ( AxesGroup.SystemData.WorkAreasMin <> 0 ) AND ( NOT HasWarning )  
THEN
  SetWarning( WarningID := RobotLibraryWarningIdEnum.WARN_FRAME_DATA_ARRAY_NOT_START_AT_ZERO, Overwrite := FALSE);
END_IF


// Check configuration parameter changed ? 
CheckParameterChanged(AxesGroup := AxesGroup);
END_METHOD

METHOD OnExecRun : DINT
VAR_IN_OUT
  /// Robot assignment of function
  AxesGroup         : AxesGroup;
END_VAR
// building rising and falling edges
_enable_R( CLK := Enable);
_enable_F( CLK := Enable);

IF ( _enable_F.Q)
THEN
  Reset(AxesGroup := AxesGroup);
END_IF


OnExecRun := RobotLibraryConstants.RUNNING;

CASE _stepCmd OF
  
  00:  IF ( _enable_R.Q )
       THEN
         // Create log entry
         CreateLogMessage ( Timestamp   := SystemTime,
                            MessageType := MessageType.CMD,
                            Severity    := Severity.INFO,
                            MessageCode := 0,
                            MessageText := 'Robot Task Enabled');
       
         // reset the rising edge
        _enable_R();
         // set busy flag
         Busy := TRUE;
         // set timeout
         SetTimeout(PT := _timeoutCmd, rTimer := _timerCmd);
         // Reset FastStop       
         AxesGroup.Cyclic.PlcToRob.FastStop := 0;
         // Reset Active command register
         AxesGroup.Acyclic.ActiveCommandRegister.Reset();
         // ST-FIX F23: the RC is still initialized from the previous enable (ACR, SEQ/ACK)
         // -> reset the interface on the RC as well
         _restartReset := AxesGroup.Cyclic.RobToPlc.TelegramState = TelegramState.INITIALIZED;
         IF ( _restartReset )
         THEN
           AxesGroup.Cyclic.PlcToRob.Control := ControlHalfByte.RESET;
         END_IF
       
         // check parameter valid
         IF ( CheckParameterValid(AxesGroup := AxesGroup) )
         THEN
           // take configuration parameter if not yet enabled
          _parCfg := ParCfg;
          // ST-FIX F103: number of telegram sequences of this configuration (not of the previous enable)
          IF ( _parCfg.Com.TwoSequences )
          THEN
            AxesGroup.State.SequenceCountSend := 1;
          ELSE
            AxesGroup.State.SequenceCountSend := 0;
          END_IF
          // ST-FIX F79: no error state of the RC seen yet in this initialization
          _initErrorState := TelegramState.UNDEFINED;
           // inc step counter
          _stepCmd := _stepCmd + 1; 
         END_IF
       END_IF
     
  01:  // ST-FIX F153: INITIALIZED without a request of this RobotTask: the RC is still
// initialized from an earlier connection -> reset the interface on the RC first
IF (( AxesGroup.Cyclic.RobToPlc.TelegramState = TelegramState.INITIALIZED ) AND
    ( AxesGroup.Cyclic.PlcToRob.Control       = ControlHalfByte.NONE      ) AND
    ( NOT _restartReset                                                   ))
THEN
  AxesGroup.Cyclic.PlcToRob.Control := ControlHalfByte.RESET;
  _restartReset := TRUE;
END_IF

